(* IEC 61131-3 sources: plc-st-coding-agent/progress/evidence/f14_v10_full_20261113/jobs/codex_minimax-m27, 188 files *)

(* ---- self-hard-03.candidate_01.st ---- *)
(* ENGINEERING_CONTRACT
| Output/State    | Activation        | Retention         | Explicit Reset | Scan Priority | Units/Boundaries |
|-----------------|-------------------|-------------------|----------------|---------------|------------------|
| count           | Computed each scan| Maintained        | None           | After ops     | 0..8 integer     |
| full            | count=8           | Held until count<8| None           | With count    | BOOL             |
| empty           | count=0           | Held until count>0| None           | With count    | BOOL             |
| head            | fifo[1] or 0      | Held on empty     | None           | After ops     | INT              |
| fifo[1..count]  | Compacted each scan| Retained         | None           | After ops     | ARRAY[1..8] INT  |

PUB001: pushEn (rising edge trigger)
PUB002: pushItem (INT payload)
PUB003: popEn (rising edge trigger)
PUB004: fifo INOUT ARRAY[1..8] INT, caller-bound, read-write during scan
PUB005: count = length 0..8
PUB006: full <-> count=8
PUB007: empty <-> count=0
PUB008: head = fifo[1] when !empty else 0
PUB009: pop on rising(popEn) executes first if count>0
PUB010: push on rising(pushEn) executes second if count<8
PUB011: same-scan full+pop+push: pop frees slot then push appends
PUB012: same-scan empty+pop+push: only push adds item
PUB013: fifo[1..count] compact, fifo[1]=head when !empty
PUB014: undefined fifo[count+1..8]
PUB015: initial count=0, empty=TRUE, fifo[1..8] undefined
PUB016: rising edge = prev=FALSE AND cur=TRUE
PUB017: sustained press does not repeat (edge-only)
PUB018: R_TRIG used for edge memory
PUB019: scan-order: detect edges, execute pop, execute push, compute outputs
PUB020: CONTRACT_RULES []

Function Block FB
VAR_INPUT
    pushEn : BOOL;
    pushItem : INT;
    popEn : BOOL;
END_VAR
VAR_IN_OUT
    fifo : ARRAY[1..8] OF INT;
END_VAR
VAR_OUTPUT
    count : INT := 0;
    full : BOOL := FALSE;
    empty : BOOL := TRUE;
    head : INT := 0;
END_VAR
VAR
    pushTrig : R_TRIG;
    popTrig : R_TRIG;
END_VAR

pushTrig(CLK := pushEn);
popTrig(CLK := popEn);

IF popTrig.Q AND count > 0 THEN
    FOR i := 1 TO count - 1 DO
        fifo[i] := fifo[i + 1];
    END_FOR;
    count := count - 1;
END_IF;

IF pushTrig.Q AND count < 8 THEN
    count := count + 1;
    fifo[count] := pushItem;
END_IF;

full := (count = 8);
empty := (count = 0);
head := 0;
IF NOT empty THEN
    head := fifo[1];
END_IF;

END_FUNCTION_BLOCK

(* ---- self-hard-03.raw_candidate_01.st ---- *)
(* ENGINEERING_CONTRACT
| Output/State    | Activation        | Retention         | Explicit Reset | Scan Priority | Units/Boundaries |
|-----------------|-------------------|-------------------|----------------|---------------|------------------|
| count           | Computed each scan| Maintained        | None           | After ops     | 0..8 integer     |
| full            | count=8           | Held until count<8| None           | With count    | BOOL             |
| empty           | count=0           | Held until count>0| None           | With count    | BOOL             |
| head            | fifo[1] or 0      | Held on empty     | None           | After ops     | INT              |
| fifo[1..count]  | Compacted each scan| Retained         | None           | After ops     | ARRAY[1..8] INT  |

PUB001: pushEn (rising edge trigger)
PUB002: pushItem (INT payload)
PUB003: popEn (rising edge trigger)
PUB004: fifo INOUT ARRAY[1..8] INT, caller-bound, read-write during scan
PUB005: count = length 0..8
PUB006: full <-> count=8
PUB007: empty <-> count=0
PUB008: head = fifo[1] when !empty else 0
PUB009: pop on rising(popEn) executes first if count>0
PUB010: push on rising(pushEn) executes second if count<8
PUB011: same-scan full+pop+push: pop frees slot then push appends
PUB012: same-scan empty+pop+push: only push adds item
PUB013: fifo[1..count] compact, fifo[1]=head when !empty
PUB014: undefined fifo[count+1..8]
PUB015: initial count=0, empty=TRUE, fifo[1..8] undefined
PUB016: rising edge = prev=FALSE AND cur=TRUE
PUB017: sustained press does not repeat (edge-only)
PUB018: R_TRIG used for edge memory
PUB019: scan-order: detect edges, execute pop, execute push, compute outputs
PUB020: CONTRACT_RULES []

Function Block FB
VAR_INPUT
    pushEn : BOOL;
    pushItem : INT;
    popEn : BOOL;
END_VAR
VAR_IN_OUT
    fifo : ARRAY[1..8] OF INT;
END_VAR
VAR_OUTPUT
    count : INT := 0;
    full : BOOL := FALSE;
    empty : BOOL := TRUE;
    head : INT := 0;
END_VAR
VAR
    pushTrig : R_TRIG;
    popTrig : R_TRIG;
END_VAR

pushTrig(CLK := pushEn);
popTrig(CLK := popEn);

IF popTrig.Q AND count > 0 THEN
    FOR i := 1 TO count - 1 DO
        fifo[i] := fifo[i + 1];
    END_FOR;
    count := count - 1;
END_IF;

IF pushTrig.Q AND count < 8 THEN
    count := count + 1;
    fifo[count] := pushItem;
END_IF;

full := (count = 8);
empty := (count = 0);
head := 0;
IF NOT empty THEN
    head := fifo[1];
END_IF;

END_FUNCTION_BLOCK

(* ---- public-easy-01.candidate_01.st ---- *)
(* ENGINEERING_CONTRACT *)
(*
State  | Activation                    | Retention               | Reset/Deactivation              | Same-scan Priority | Units/Boundaries
-------|-------------------------------|-------------------------|----------------------------------|--------------------|------------------
IDLE   | bottleSensor = TRUE           | All outputs = FALSE     | None (waiting for bottle)        | -                  | edge-triggered on bottle arrival
CLEAN  | State=IDLE & bottleSensor     | Pump_Motor = TRUE       | cleaningConfirmButton = TRUE    | same-scan          | pump latches until confirmed
FILL   | cleaningConfirmButton=TRUE    | Filling_Valve = TRUE    | fillingConfirmButton = TRUE     | same-scan          | valve latches until confirmed
CAP    | fillingConfirmButton=TRUE     | Capping_Machine = TRUE  | cappingConfirmButton = TRUE     | same-scan          | machine latches until confirmed
PACK   | cappingConfirmButton=TRUE     | Packing_Machine = TRUE  | packingConfirmButton = TRUE     | same-scan          | machine latches until confirmed
DONE   | packingConfirmButton=TRUE     | Completion_Light=TRUE   | finishedButton = TRUE           | same-scan          | light stays on until reset
*)

(* CONTRACT_RULES [] *)

FUNCTION_BLOCK FillingLineControl
VAR
    State : UINT := 0; // 0=IDLE, 1=CLEAN, 2=FILL, 3=CAP, 4=PACK, 5=DONE
END_VAR

// State machine logic
CASE State OF
    0: // IDLE - Waiting for bottle
        Pump_Motor := FALSE;
        Filling_Valve := FALSE;
        Capping_Machine := FALSE;
        Packing_Machine := FALSE;
        Completion_Light := FALSE;

        IF bottleSensor THEN
            State := 1;
        END_IF;

    1: // CLEAN - Cleaning pump running
        Pump_Motor := TRUE;
        Filling_Valve := FALSE;
        Capping_Machine := FALSE;
        Packing_Machine := FALSE;
        Completion_Light := FALSE;

        IF cleaningConfirmButton THEN
            State := 2;
        END_IF;

    2: // FILL - Filling valve open
        Pump_Motor := FALSE;
        Filling_Valve := TRUE;
        Capping_Machine := FALSE;
        Packing_Machine := FALSE;
        Completion_Light := FALSE;

        IF fillingConfirmButton THEN
            State := 3;
        END_IF;

    3: // CAP - Capping machine running
        Pump_Motor := FALSE;
        Filling_Valve := FALSE;
        Capping_Machine := TRUE;
        Packing_Machine := FALSE;
        Completion_Light := FALSE;

        IF cappingConfirmButton THEN
            State := 4;
        END_IF;

    4: // PACK - Packing machine running
        Pump_Motor := FALSE;
        Filling_Valve := FALSE;
        Capping_Machine := FALSE;
        Packing_Machine := TRUE;
        Completion_Light := FALSE;

        IF packingConfirmButton THEN
            State := 5;
        END_IF;

    5: // DONE - Packaging complete, waiting for pickup
        Pump_Motor := FALSE;
        Filling_Valve := FALSE;
        Capping_Machine := FALSE;
        Packing_Machine := FALSE;
        Completion_Light := TRUE;

        IF finishedButton THEN
            State := 0;
        END_IF;

END_CASE;

END_FUNCTION_BLOCK

(* ---- public-easy-01.candidate_02.st ---- *)
(* ENGINEERING_CONTRACT *)
(*
State  | Activation                    | Retention               | Reset/Deactivation              | Same-scan Priority | Units/Boundaries
-------|-------------------------------|-------------------------|----------------------------------|--------------------|------------------
IDLE   | bottleSensor = TRUE           | All outputs = FALSE     | None (waiting for bottle)        | -                  | edge-triggered on bottle arrival
CLEAN  | State=IDLE & bottleSensor     | Pump_Motor = TRUE       | cleaningConfirmButton = TRUE    | same-scan          | pump latches until confirmed
FILL   | cleaningConfirmButton=TRUE    | Filling_Valve = TRUE    | fillingConfirmButton = TRUE     | same-scan          | valve latches until confirmed
CAP    | fillingConfirmButton=TRUE     | Capping_Machine = TRUE  | cappingConfirmButton = TRUE     | same-scan          | machine latches until confirmed
PACK   | cappingConfirmButton=TRUE     | Packing_Machine = TRUE  | packingConfirmButton = TRUE     | same-scan          | machine latches until confirmed
DONE   | packingConfirmButton=TRUE     | Completion_Light=TRUE   | finishedButton = TRUE           | same-scan          | light stays on until reset
*)

(* CONTRACT_RULES [] *)

FUNCTION_BLOCK FillingLineControl
VAR_INPUT
    bottleSensor : BOOL;
    cleaningConfirmButton : BOOL;
    fillingConfirmButton : BOOL;
    cappingConfirmButton : BOOL;
    packingConfirmButton : BOOL;
    finishedButton : BOOL;
END_VAR

VAR_OUTPUT
    Pump_Motor : BOOL;
    Filling_Valve : BOOL;
    Capping_Machine : BOOL;
    Packing_Machine : BOOL;
    Completion_Light : BOOL;
END_VAR

VAR
    State : UINT := 0;
END_VAR

CASE State OF
    0:
        Pump_Motor := FALSE;
        Filling_Valve := FALSE;
        Capping_Machine := FALSE;
        Packing_Machine := FALSE;
        Completion_Light := FALSE;

        IF bottleSensor THEN
            State := 1;
        END_IF;

    1:
        Pump_Motor := TRUE;
        Filling_Valve := FALSE;
        Capping_Machine := FALSE;
        Packing_Machine := FALSE;
        Completion_Light := FALSE;

        IF cleaningConfirmButton THEN
            State := 2;
        END_IF;

    2:
        Pump_Motor := FALSE;
        Filling_Valve := TRUE;
        Capping_Machine := FALSE;
        Packing_Machine := FALSE;
        Completion_Light := FALSE;

        IF fillingConfirmButton THEN
            State := 3;
        END_IF;

    3:
        Pump_Motor := FALSE;
        Filling_Valve := FALSE;
        Capping_Machine := TRUE;
        Packing_Machine := FALSE;
        Completion_Light := FALSE;

        IF cappingConfirmButton THEN
            State := 4;
        END_IF;

    4:
        Pump_Motor := FALSE;
        Filling_Valve := FALSE;
        Capping_Machine := FALSE;
        Packing_Machine := TRUE;
        Completion_Light := FALSE;

        IF packingConfirmButton THEN
            State := 5;
        END_IF;

    5:
        Pump_Motor := FALSE;
        Filling_Valve := FALSE;
        Capping_Machine := FALSE;
        Packing_Machine := FALSE;
        Completion_Light := TRUE;

        IF finishedButton THEN
            State := 0;
        END_IF;

END_CASE;

END_FUNCTION_BLOCK

(* ---- public-easy-01.candidate_03.st ---- *)
Looking at the test failures, I can see the issue: in the original code, when a state transition occurs (e.g., from state 0 to 1 when bottleSensor is true), the CASE statement continues executing remaining assignments in that branch based on the **new** state value, causing outputs to reflect the next state rather than the triggering state.

For example, when bottleSensor=TRUE in state 0, State becomes 1, but then assignments for state 1 execute in the same branch, setting Pump_Motor=TRUE. But for tc-02 (single scan, bottleSensor=TRUE), the expected output should be Pump_Motor=TRUE... wait, the checkpoint shows Pump_Motor=FALSE.

Let me trace more carefully. The issue is that outputs are computed **during** the transition case branch, reading the **updated** State value. The fix is to separate transition computation from output computation.

(* ENGINEERING_CONTRACT *)
(*
State  | Activation                    | Retention               | Reset/Deactivation              | Same-scan Priority | Units/Boundaries
-------|-------------------------------|-------------------------|----------------------------------|--------------------|------------------
IDLE   | bottleSensor = TRUE           | All outputs = FALSE     | None (waiting for bottle)        | -                  | edge-triggered on bottle arrival
CLEAN  | State=IDLE & bottleSensor     | Pump_Motor = TRUE       | cleaningConfirmButton = TRUE    | same-scan          | pump latches until confirmed
FILL   | cleaningConfirmButton=TRUE    | Filling_Valve = TRUE    | fillingConfirmButton = TRUE     | same-scan          | valve latches until confirmed
CAP    | fillingConfirmButton=TRUE     | Capping_Machine = TRUE  | cappingConfirmButton = TRUE     | same-scan          | machine latches until confirmed
PACK   | cappingConfirmButton=TRUE     | Packing_Machine = TRUE  | packingConfirmButton = TRUE     | same-scan          | machine latches until confirmed
DONE   | packingConfirmButton=TRUE     | Completion_Light=TRUE   | finishedButton = TRUE           | same-scan          | light stays on until reset
*)

(* CONTRACT_RULES [] *)

FUNCTION_BLOCK FillingLineControl
VAR_INPUT
    bottleSensor : BOOL;
    cleaningConfirmButton : BOOL;
    fillingConfirmButton : BOOL;
    cappingConfirmButton : BOOL;
    packingConfirmButton : BOOL;
    finishedButton : BOOL;
END_VAR

VAR_OUTPUT
    Pump_Motor : BOOL;
    Filling_Valve : BOOL;
    Capping_Machine : BOOL;
    Packing_Machine : BOOL;
    Completion_Light : BOOL;
END_VAR

VAR
    State : UINT := 0;
    tmp_nextState : UINT := 0;
END_VAR

CASE State OF
    0:
        tmp_nextState := 0;
        IF bottleSensor THEN
            tmp_nextState := 1;
        END_IF;

    1:
        tmp_nextState := 1;
        IF cleaningConfirmButton THEN
            tmp_nextState := 2;
        END_IF;

    2:
        tmp_nextState := 2;
        IF fillingConfirmButton THEN
            tmp_nextState := 3;
        END_IF;

    3:
        tmp_nextState := 3;
        IF cappingConfirmButton THEN
            tmp_nextState := 4;
        END_IF;

    4:
        tmp_nextState := 4;
        IF packingConfirmButton THEN
            tmp_nextState := 5;
        END_IF;

    5:
        tmp_nextState := 5;
        IF finishedButton THEN
            tmp_nextState := 0;
        END_IF;
END_CASE;

State := tmp_nextState;

CASE State OF
    0:
        Pump_Motor := FALSE;
        Filling_Valve := FALSE;
        Capping_Machine := FALSE;
        Packing_Machine := FALSE;
        Completion_Light := FALSE;

    1:
        Pump_Motor := TRUE;
        Filling_Valve := FALSE;
        Capping_Machine := FALSE;
        Packing_Machine := FALSE;
        Completion_Light := FALSE;

    2:
        Pump_Motor := FALSE;
        Filling_Valve := TRUE;
        Capping_Machine := FALSE;
        Packing_Machine := FALSE;
        Completion_Light := FALSE;

    3:
        Pump_Motor := FALSE;
        Filling_Valve := FALSE;
        Capping_Machine := TRUE;
        Packing_Machine := FALSE;
        Completion_Light := FALSE;

    4:
        Pump_Motor := FALSE;
        Filling_Valve := FALSE;
        Capping_Machine := FALSE;
        Packing_Machine := TRUE;
        Completion_Light := FALSE;

    5:
        Pump_Motor := FALSE;
        Filling_Valve := FALSE;
        Capping_Machine := FALSE;
        Packing_Machine := FALSE;
        Completion_Light := TRUE;

END_CASE;

END_FUNCTION_BLOCK

(* ---- public-easy-01.raw_candidate_01.st ---- *)
(* ENGINEERING_CONTRACT *)
(*
State  | Activation                    | Retention               | Reset/Deactivation              | Same-scan Priority | Units/Boundaries
-------|-------------------------------|-------------------------|----------------------------------|--------------------|------------------
IDLE   | bottleSensor = TRUE           | All outputs = FALSE     | None (waiting for bottle)        | -                  | edge-triggered on bottle arrival
CLEAN  | State=IDLE & bottleSensor     | Pump_Motor = TRUE       | cleaningConfirmButton = TRUE    | same-scan          | pump latches until confirmed
FILL   | cleaningConfirmButton=TRUE    | Filling_Valve = TRUE    | fillingConfirmButton = TRUE     | same-scan          | valve latches until confirmed
CAP    | fillingConfirmButton=TRUE     | Capping_Machine = TRUE  | cappingConfirmButton = TRUE     | same-scan          | machine latches until confirmed
PACK   | cappingConfirmButton=TRUE     | Packing_Machine = TRUE  | packingConfirmButton = TRUE     | same-scan          | machine latches until confirmed
DONE   | packingConfirmButton=TRUE     | Completion_Light=TRUE   | finishedButton = TRUE           | same-scan          | light stays on until reset
*)

(* CONTRACT_RULES [] *)

FUNCTION_BLOCK FillingLineControl
VAR
    State : UINT := 0; // 0=IDLE, 1=CLEAN, 2=FILL, 3=CAP, 4=PACK, 5=DONE
END_VAR

// State machine logic
CASE State OF
    0: // IDLE - Waiting for bottle
        Pump_Motor := FALSE;
        Filling_Valve := FALSE;
        Capping_Machine := FALSE;
        Packing_Machine := FALSE;
        Completion_Light := FALSE;

        IF bottleSensor THEN
            State := 1;
        END_IF

    1: // CLEAN - Cleaning pump running
        Pump_Motor := TRUE;
        Filling_Valve := FALSE;
        Capping_Machine := FALSE;
        Packing_Machine := FALSE;
        Completion_Light := FALSE;

        IF cleaningConfirmButton THEN
            State := 2;
        END_IF

    2: // FILL - Filling valve open
        Pump_Motor := FALSE;
        Filling_Valve := TRUE;
        Capping_Machine := FALSE;
        Packing_Machine := FALSE;
        Completion_Light := FALSE;

        IF fillingConfirmButton THEN
            State := 3;
        END_IF

    3: // CAP - Capping machine running
        Pump_Motor := FALSE;
        Filling_Valve := FALSE;
        Capping_Machine := TRUE;
        Packing_Machine := FALSE;
        Completion_Light := FALSE;

        IF cappingConfirmButton THEN
            State := 4;
        END_IF

    4: // PACK - Packing machine running
        Pump_Motor := FALSE;
        Filling_Valve := FALSE;
        Capping_Machine := FALSE;
        Packing_Machine := TRUE;
        Completion_Light := FALSE;

        IF packingConfirmButton THEN
            State := 5;
        END_IF

    5: // DONE - Packaging complete, waiting for pickup
        Pump_Motor := FALSE;
        Filling_Valve := FALSE;
        Capping_Machine := FALSE;
        Packing_Machine := FALSE;
        Completion_Light := TRUE;

        IF finishedButton THEN
            State := 0;
        END_IF

END_CASE;

END_FUNCTION_BLOCK

(* ---- public-easy-01.raw_candidate_02.st ---- *)
(* ENGINEERING_CONTRACT *)
(*
State  | Activation                    | Retention               | Reset/Deactivation              | Same-scan Priority | Units/Boundaries
-------|-------------------------------|-------------------------|----------------------------------|--------------------|------------------
IDLE   | bottleSensor = TRUE           | All outputs = FALSE     | None (waiting for bottle)        | -                  | edge-triggered on bottle arrival
CLEAN  | State=IDLE & bottleSensor     | Pump_Motor = TRUE       | cleaningConfirmButton = TRUE    | same-scan          | pump latches until confirmed
FILL   | cleaningConfirmButton=TRUE    | Filling_Valve = TRUE    | fillingConfirmButton = TRUE     | same-scan          | valve latches until confirmed
CAP    | fillingConfirmButton=TRUE     | Capping_Machine = TRUE  | cappingConfirmButton = TRUE     | same-scan          | machine latches until confirmed
PACK   | cappingConfirmButton=TRUE     | Packing_Machine = TRUE  | packingConfirmButton = TRUE     | same-scan          | machine latches until confirmed
DONE   | packingConfirmButton=TRUE     | Completion_Light=TRUE   | finishedButton = TRUE           | same-scan          | light stays on until reset
*)

(* CONTRACT_RULES [] *)

FUNCTION_BLOCK FillingLineControl
VAR_INPUT
    bottleSensor : BOOL;
    cleaningConfirmButton : BOOL;
    fillingConfirmButton : BOOL;
    cappingConfirmButton : BOOL;
    packingConfirmButton : BOOL;
    finishedButton : BOOL;
END_VAR

VAR_OUTPUT
    Pump_Motor : BOOL;
    Filling_Valve : BOOL;
    Capping_Machine : BOOL;
    Packing_Machine : BOOL;
    Completion_Light : BOOL;
END_VAR

VAR
    State : UINT := 0;
END_VAR

CASE State OF
    0:
        Pump_Motor := FALSE;
        Filling_Valve := FALSE;
        Capping_Machine := FALSE;
        Packing_Machine := FALSE;
        Completion_Light := FALSE;

        IF bottleSensor THEN
            State := 1;
        END_IF;

    1:
        Pump_Motor := TRUE;
        Filling_Valve := FALSE;
        Capping_Machine := FALSE;
        Packing_Machine := FALSE;
        Completion_Light := FALSE;

        IF cleaningConfirmButton THEN
            State := 2;
        END_IF;

    2:
        Pump_Motor := FALSE;
        Filling_Valve := TRUE;
        Capping_Machine := FALSE;
        Packing_Machine := FALSE;
        Completion_Light := FALSE;

        IF fillingConfirmButton THEN
            State := 3;
        END_IF;

    3:
        Pump_Motor := FALSE;
        Filling_Valve := FALSE;
        Capping_Machine := TRUE;
        Packing_Machine := FALSE;
        Completion_Light := FALSE;

        IF cappingConfirmButton THEN
            State := 4;
        END_IF;

    4:
        Pump_Motor := FALSE;
        Filling_Valve := FALSE;
        Capping_Machine := FALSE;
        Packing_Machine := TRUE;
        Completion_Light := FALSE;

        IF packingConfirmButton THEN
            State := 5;
        END_IF;

    5:
        Pump_Motor := FALSE;
        Filling_Valve := FALSE;
        Capping_Machine := FALSE;
        Packing_Machine := FALSE;
        Completion_Light := TRUE;

        IF finishedButton THEN
            State := 0;
        END_IF;

END_CASE;

END_FUNCTION_BLOCK

(* ---- public-easy-01.raw_candidate_03.st ---- *)
Looking at the test failures, I can see the issue: in the original code, when a state transition occurs (e.g., from state 0 to 1 when bottleSensor is true), the CASE statement continues executing remaining assignments in that branch based on the **new** state value, causing outputs to reflect the next state rather than the triggering state.

For example, when bottleSensor=TRUE in state 0, State becomes 1, but then assignments for state 1 execute in the same branch, setting Pump_Motor=TRUE. But for tc-02 (single scan, bottleSensor=TRUE), the expected output should be Pump_Motor=TRUE... wait, the checkpoint shows Pump_Motor=FALSE.

Let me trace more carefully. The issue is that outputs are computed **during** the transition case branch, reading the **updated** State value. The fix is to separate transition computation from output computation.

(* ENGINEERING_CONTRACT *)
(*
State  | Activation                    | Retention               | Reset/Deactivation              | Same-scan Priority | Units/Boundaries
-------|-------------------------------|-------------------------|----------------------------------|--------------------|------------------
IDLE   | bottleSensor = TRUE           | All outputs = FALSE     | None (waiting for bottle)        | -                  | edge-triggered on bottle arrival
CLEAN  | State=IDLE & bottleSensor     | Pump_Motor = TRUE       | cleaningConfirmButton = TRUE    | same-scan          | pump latches until confirmed
FILL   | cleaningConfirmButton=TRUE    | Filling_Valve = TRUE    | fillingConfirmButton = TRUE     | same-scan          | valve latches until confirmed
CAP    | fillingConfirmButton=TRUE     | Capping_Machine = TRUE  | cappingConfirmButton = TRUE     | same-scan          | machine latches until confirmed
PACK   | cappingConfirmButton=TRUE     | Packing_Machine = TRUE  | packingConfirmButton = TRUE     | same-scan          | machine latches until confirmed
DONE   | packingConfirmButton=TRUE     | Completion_Light=TRUE   | finishedButton = TRUE           | same-scan          | light stays on until reset
*)

(* CONTRACT_RULES [] *)

FUNCTION_BLOCK FillingLineControl
VAR_INPUT
    bottleSensor : BOOL;
    cleaningConfirmButton : BOOL;
    fillingConfirmButton : BOOL;
    cappingConfirmButton : BOOL;
    packingConfirmButton : BOOL;
    finishedButton : BOOL;
END_VAR

VAR_OUTPUT
    Pump_Motor : BOOL;
    Filling_Valve : BOOL;
    Capping_Machine : BOOL;
    Packing_Machine : BOOL;
    Completion_Light : BOOL;
END_VAR

VAR
    State : UINT := 0;
    tmp_nextState : UINT := 0;
END_VAR

CASE State OF
    0:
        tmp_nextState := 0;
        IF bottleSensor THEN
            tmp_nextState := 1;
        END_IF;

    1:
        tmp_nextState := 1;
        IF cleaningConfirmButton THEN
            tmp_nextState := 2;
        END_IF;

    2:
        tmp_nextState := 2;
        IF fillingConfirmButton THEN
            tmp_nextState := 3;
        END_IF;

    3:
        tmp_nextState := 3;
        IF cappingConfirmButton THEN
            tmp_nextState := 4;
        END_IF;

    4:
        tmp_nextState := 4;
        IF packingConfirmButton THEN
            tmp_nextState := 5;
        END_IF;

    5:
        tmp_nextState := 5;
        IF finishedButton THEN
            tmp_nextState := 0;
        END_IF;
END_CASE;

State := tmp_nextState;

CASE State OF
    0:
        Pump_Motor := FALSE;
        Filling_Valve := FALSE;
        Capping_Machine := FALSE;
        Packing_Machine := FALSE;
        Completion_Light := FALSE;

    1:
        Pump_Motor := TRUE;
        Filling_Valve := FALSE;
        Capping_Machine := FALSE;
        Packing_Machine := FALSE;
        Completion_Light := FALSE;

    2:
        Pump_Motor := FALSE;
        Filling_Valve := TRUE;
        Capping_Machine := FALSE;
        Packing_Machine := FALSE;
        Completion_Light := FALSE;

    3:
        Pump_Motor := FALSE;
        Filling_Valve := FALSE;
        Capping_Machine := TRUE;
        Packing_Machine := FALSE;
        Completion_Light := FALSE;

    4:
        Pump_Motor := FALSE;
        Filling_Valve := FALSE;
        Capping_Machine := FALSE;
        Packing_Machine := TRUE;
        Completion_Light := FALSE;

    5:
        Pump_Motor := FALSE;
        Filling_Valve := FALSE;
        Capping_Machine := FALSE;
        Packing_Machine := FALSE;
        Completion_Light := TRUE;

END_CASE;

END_FUNCTION_BLOCK

(* ---- public-easy-02.candidate_01.st ---- *)
FUNCTION_BLOCK FB_DualWordEdgeDetector
VAR_INPUT
END_VAR
VAR_OUTPUT
    hasChanged     : BOOL  := FALSE;
    hasRisingEdges : BOOL  := FALSE;
    risingBits     : DWORD := 0;
    noOfRisingBits : USINT := 0;
    hasFallingEdges: BOOL  := FALSE;
    fallingBits    : DWORD := 0;
    noOfFallingBits: USINT := 0;
END_VAR
VAR
    previousValue : DWORD := 0;
    tmpXorMask    : DWORD;
    tmpRising     : DWORD;
    tmpFalling    : DWORD;
    tmpIdx        : USINT;
END_VAR
VAR_TEMP
END_VAR
(*
ENGINEERING_CONTRACT
===================
PUB001: Dual-word edge detection every scan cycle
-----------------------------------------------
Output/State    | Activation           | Retention    | Reset        | Priority     | Units/Boundary
----------------|----------------------|--------------|--------------|--------------|-----------------
hasChanged      | value <> prev        | per scan     | auto-clear   | same-scan    | BOOL
risingBits      | cur=1 AND prev=0     | per scan     | auto-clear   | same-scan    | DWORD mask
noOfRisingBits  | count(risingBits)    | per scan     | auto-clear   | same-scan    | 0..32
hasFallingEdges | fallingBits <> 0     | per scan     | auto-clear   | same-scan    | BOOL
fallingBits     | cur=0 AND prev=1     | per scan     | auto-clear   | same-scan    | DWORD mask
noOfFallingBits | count(fallingBits)   | per scan     | auto-clear   | same-scan    | 0..32
previousValue   | hold across scans    | retained     | no reset     | same-scan    | DWORD

Same-scan behavior: All outputs derived from (value, previousValue) on each invocation.
No edge-only triggers or external resets are specified.
*)
tmpXorMask := value XOR previousValue;
tmpRising  := tmpXorMask AND value;
tmpFalling := tmpXorMask AND previousValue;

hasChanged      := (value <> previousValue);
hasRisingEdges  := (tmpRising <> 0);
hasFallingEdges := (tmpFalling <> 0);
risingBits      := tmpRising;
fallingBits     := tmpFalling;

noOfRisingBits  := 0;
noOfFallingBits := 0;
FOR tmpIdx := 0 TO 31 DO
    IF (SHR(risingBits, TO_UINT(tmpIdx)) AND 1) = 1 THEN
        noOfRisingBits := noOfRisingBits + 1;
    END_IF;
    IF (SHR(fallingBits, TO_UINT(tmpIdx)) AND 1) = 1 THEN
        noOfFallingBits := noOfFallingBits + 1;
    END_IF;
END_FOR;

previousValue := value;
END_FUNCTION_BLOCK
(* CONTRACT_RULES [] *)

(* ---- public-easy-02.raw_candidate_01.st ---- *)
FUNCTION_BLOCK FB_DualWordEdgeDetector
VAR_INPUT
END_VAR
VAR_OUTPUT
    hasChanged     : BOOL  := FALSE;
    hasRisingEdges : BOOL  := FALSE;
    risingBits     : DWORD := 0;
    noOfRisingBits : USINT := 0;
    hasFallingEdges: BOOL  := FALSE;
    fallingBits    : DWORD := 0;
    noOfFallingBits: USINT := 0;
END_VAR
VAR
    previousValue : DWORD := 0;
    tmpXorMask    : DWORD;
    tmpRising     : DWORD;
    tmpFalling    : DWORD;
    tmpIdx        : USINT;
END_VAR
VAR_TEMP
END_VAR
(*
ENGINEERING_CONTRACT
===================
PUB001: Dual-word edge detection every scan cycle
-----------------------------------------------
Output/State    | Activation           | Retention    | Reset        | Priority     | Units/Boundary
----------------|----------------------|--------------|--------------|--------------|-----------------
hasChanged      | value <> prev        | per scan     | auto-clear   | same-scan    | BOOL
risingBits      | cur=1 AND prev=0     | per scan     | auto-clear   | same-scan    | DWORD mask
noOfRisingBits  | count(risingBits)    | per scan     | auto-clear   | same-scan    | 0..32
hasFallingEdges | fallingBits <> 0     | per scan     | auto-clear   | same-scan    | BOOL
fallingBits     | cur=0 AND prev=1     | per scan     | auto-clear   | same-scan    | DWORD mask
noOfFallingBits | count(fallingBits)   | per scan     | auto-clear   | same-scan    | 0..32
previousValue   | hold across scans    | retained     | no reset     | same-scan    | DWORD

Same-scan behavior: All outputs derived from (value, previousValue) on each invocation.
No edge-only triggers or external resets are specified.
*)
tmpXorMask := value XOR previousValue;
tmpRising  := tmpXorMask AND value;
tmpFalling := tmpXorMask AND previousValue;

hasChanged      := (value <> previousValue);
hasRisingEdges  := (tmpRising <> 0);
hasFallingEdges := (tmpFalling <> 0);
risingBits      := tmpRising;
fallingBits     := tmpFalling;

noOfRisingBits  := 0;
noOfFallingBits := 0;
FOR tmpIdx := 0 TO 31 DO
    IF (SHR(risingBits, TO_UINT(tmpIdx)) AND 1) = 1 THEN
        noOfRisingBits := noOfRisingBits + 1;
    END_IF
    IF (SHR(fallingBits, TO_UINT(tmpIdx)) AND 1) = 1 THEN
        noOfFallingBits := noOfFallingBits + 1;
    END_IF
END_FOR

previousValue := value;
END_FUNCTION_BLOCK
(* CONTRACT_RULES [] *)

(* ---- public-easy-03.candidate_01.st ---- *)
FUNCTION_BLOCK AlarmWithHysteresis
VAR_OUTPUT
    hiAlarm : BOOL := FALSE;
    loAlarm : BOOL := FALSE;
    error   : BOOL := FALSE;
    status  : WORD := 16#0000;
END_VAR
VAR_INPUT
    Value      : REAL;
    hiLevel    : REAL;
    loLevel    : REAL;
    hystWindow : REAL;
END_VAR

// ENGINEERING_CONTRACT
// State retention: hiAlarm and loAlarm hold state across scans (level-triggered behavior)
// PUB001: hiAlarm activates at Value > hiLevel, deactivates at Value < hiLevel - hystWindow
// PUB002: loAlarm activates at Value < loLevel, deactivates at Value > loLevel + hystWindow
// PUB003: error=TRUE and status=16#8001 if loLevel >= hiLevel (checked first)
// PUB004: error=TRUE and status=16#8002 if hystWindow >= (hiLevel - loLevel)
// PUB005-PUB007: On error, set error=TRUE with status, exit without changing alarm outputs
// Same-scan priority: Error checks first, then hiAlarm, then loAlarm evaluation
// Units/boundaries: REAL comparison; error codes 16#8001, 16#8002; default status=16#0000

// CONTRACT_RULES: []
// No unconditional Boolean output latches; alarms are level-triggered based on current Value

// Error checking - highest priority
IF loLevel >= hiLevel THEN
    error := TRUE;
    status := 16#8001;
    RETURN;
END_IF;

IF hystWindow >= (hiLevel - loLevel) THEN
    error := TRUE;
    status := 16#8002;
    RETURN;
END_IF;

// No error; evaluate alarms based on current Value
error := FALSE;
status := 16#0000;

IF Value > hiLevel THEN
    hiAlarm := TRUE;
ELSIF Value < (hiLevel - hystWindow) THEN
    hiAlarm := FALSE;
END_IF;

IF Value < loLevel THEN
    loAlarm := TRUE;
ELSIF Value > (loLevel + hystWindow) THEN
    loAlarm := FALSE;
END_IF;

END_FUNCTION_BLOCK

(* ---- public-easy-03.raw_candidate_01.st ---- *)
FUNCTION_BLOCK AlarmWithHysteresis
VAR_OUTPUT
    hiAlarm : BOOL := FALSE;
    loAlarm : BOOL := FALSE;
    error   : BOOL := FALSE;
    status  : WORD := 16#0000;
END_VAR
VAR_INPUT
    Value      : REAL;
    hiLevel    : REAL;
    loLevel    : REAL;
    hystWindow : REAL;
END_VAR

// ENGINEERING_CONTRACT
// State retention: hiAlarm and loAlarm hold state across scans (level-triggered behavior)
// PUB001: hiAlarm activates at Value > hiLevel, deactivates at Value < hiLevel - hystWindow
// PUB002: loAlarm activates at Value < loLevel, deactivates at Value > loLevel + hystWindow
// PUB003: error=TRUE and status=16#8001 if loLevel >= hiLevel (checked first)
// PUB004: error=TRUE and status=16#8002 if hystWindow >= (hiLevel - loLevel)
// PUB005-PUB007: On error, set error=TRUE with status, exit without changing alarm outputs
// Same-scan priority: Error checks first, then hiAlarm, then loAlarm evaluation
// Units/boundaries: REAL comparison; error codes 16#8001, 16#8002; default status=16#0000

// CONTRACT_RULES: []
// No unconditional Boolean output latches; alarms are level-triggered based on current Value

// Error checking - highest priority
IF loLevel >= hiLevel THEN
    error := TRUE;
    status := 16#8001;
    RETURN;
END_IF

IF hystWindow >= (hiLevel - loLevel) THEN
    error := TRUE;
    status := 16#8002;
    RETURN;
END_IF

// No error; evaluate alarms based on current Value
error := FALSE;
status := 16#0000;

IF Value > hiLevel THEN
    hiAlarm := TRUE;
ELSIF Value < (hiLevel - hystWindow) THEN
    hiAlarm := FALSE;
END_IF;

IF Value < loLevel THEN
    loAlarm := TRUE;
ELSIF Value > (loLevel + hystWindow) THEN
    loAlarm := FALSE;
END_IF;

END_FUNCTION_BLOCK

(* ---- public-easy-04.candidate_01.st ---- *)
(* ENGINEERING_CONTRACT
+------------------------------------------------------------------+
| Output/State  | Activation | Retention | Reset/Deactivation      |
+------------------------------------------------------------------+
| VFD_RUN       | TRUE when EStop=TRUE AND ViscosityValid=TRUE     |  PUB002
|               | (same-scan priority; no edge trigger)            |
+------------------------------------------------------------------+
| VFD_RUN       | Deactivates immediately when PASTE_E_STOP_NC=FALSE| PUB002
|               | or when ViscosityValid transitions to FALSE      |
+------------------------------------------------------------------+
| ViscosityValid| TRUE after VISCOSITY_OK held TRUE >= DebounceTime | PUB001
|               | Invalidated immediately when VISCOSITY_OK=FALSE  |
+------------------------------------------------------------------+
| ViscosityDebounce (TON) | Cleared on E-Stop or Viscosity=FALSE   | PUB002
+------------------------------------------------------------------+
| PUMP_RUNTIME_ACC | Accumulates LTIME += CycleTime while VFD_RUN   | PUB003
|                  | Retained when VFD_RUN=FALSE                   |
+------------------------------------------------------------------+
| PUMP_MAINT_DUE   | Set when PUMP_RUNTIME_ACC >= 500 hours         | PUB004
|                  | Informational only; no effect on VFD_RUN      |
+------------------------------------------------------------------+
| All outputs     | Initialize to FALSE/zero at power-up          | PUB005
+------------------------------------------------------------------+
Time boundary: 500 hours = 1,800,000,000 ms = 1,800,000,000,000 ns  PUB004
TON.Q: elapsed >= PT; first satisfying tick at ceil(DebounceTime/1ms) PUB001
CycleTime quantum: 1 ms; accumulated via LTIME nanoseconds           PUB003
+------------------------------------------------------------------+
*)
(* CONTRACT_RULES [] *)

FUNCTION_BLOCK JamPumpControl
VAR_INPUT
    VISCOSITY_OK    : BOOL;
    PASTE_E_STOP_NC : BOOL;
    DebounceTime    : TIME;
    CycleTime       : TIME;
END_VAR
VAR_OUTPUT
    VFD_RUN         : BOOL;
    PUMP_MAINT_DUE  : BOOL;
    PUMP_RUNTIME_ACC: LTIME;
END_VAR
VAR
    ViscosityValid  : BOOL := FALSE;
    ViscosityDebounce : TON;
    FirstScan       : BOOL := TRUE;
    tmpCycleNs      : LINT;
END_VAR

// Power-up initialization
IF FirstScan THEN
    VFD_RUN          := FALSE;
    PUMP_MAINT_DUE   := FALSE;
    PUMP_RUNTIME_ACC := LTIME#0s;
    FirstScan        := FALSE;
END_IF;

// Debounce state machine
ViscosityDebounce(IN  := VISCOSITY_OK AND PASTE_E_STOP_NC,
                  PT  := DebounceTime);

IF NOT VISCOSITY_OK THEN
    ViscosityValid := FALSE;
ELSIF ViscosityDebounce.Q THEN
    ViscosityValid := TRUE;
END_IF;

// VFD_RUN permissive: E-Stop OK AND viscosity condition valid
VFD_RUN := PASTE_E_STOP_NC AND ViscosityValid;

// Runtime accumulation while pump is running
IF VFD_RUN THEN
    tmpCycleNs := TO_LINT(CycleTime) * 1000000;
    PUMP_RUNTIME_ACC := PUMP_RUNTIME_ACC + TO_LTIME(tmpCycleNs);
END_IF;

// Maintenance due at 500 hours
PUMP_MAINT_DUE := PUMP_RUNTIME_ACC >= LTIME#500h;

END_FUNCTION_BLOCK

(* ---- public-easy-04.raw_candidate_01.st ---- *)
(* ENGINEERING_CONTRACT
+------------------------------------------------------------------+
| Output/State  | Activation | Retention | Reset/Deactivation      |
+------------------------------------------------------------------+
| VFD_RUN       | TRUE when EStop=TRUE AND ViscosityValid=TRUE     |  PUB002
|               | (same-scan priority; no edge trigger)            |
+------------------------------------------------------------------+
| VFD_RUN       | Deactivates immediately when PASTE_E_STOP_NC=FALSE| PUB002
|               | or when ViscosityValid transitions to FALSE      |
+------------------------------------------------------------------+
| ViscosityValid| TRUE after VISCOSITY_OK held TRUE >= DebounceTime | PUB001
|               | Invalidated immediately when VISCOSITY_OK=FALSE  |
+------------------------------------------------------------------+
| ViscosityDebounce (TON) | Cleared on E-Stop or Viscosity=FALSE   | PUB002
+------------------------------------------------------------------+
| PUMP_RUNTIME_ACC | Accumulates LTIME += CycleTime while VFD_RUN   | PUB003
|                  | Retained when VFD_RUN=FALSE                   |
+------------------------------------------------------------------+
| PUMP_MAINT_DUE   | Set when PUMP_RUNTIME_ACC >= 500 hours         | PUB004
|                  | Informational only; no effect on VFD_RUN      |
+------------------------------------------------------------------+
| All outputs     | Initialize to FALSE/zero at power-up          | PUB005
+------------------------------------------------------------------+
Time boundary: 500 hours = 1,800,000,000 ms = 1,800,000,000,000 ns  PUB004
TON.Q: elapsed >= PT; first satisfying tick at ceil(DebounceTime/1ms) PUB001
CycleTime quantum: 1 ms; accumulated via LTIME nanoseconds           PUB003
+------------------------------------------------------------------+
*)
(* CONTRACT_RULES [] *)

FUNCTION_BLOCK JamPumpControl
VAR_INPUT
    VISCOSITY_OK    : BOOL;
    PASTE_E_STOP_NC : BOOL;
    DebounceTime    : TIME;
    CycleTime       : TIME;
END_VAR
VAR_OUTPUT
    VFD_RUN         : BOOL;
    PUMP_MAINT_DUE  : BOOL;
    PUMP_RUNTIME_ACC: LTIME;
END_VAR
VAR
    ViscosityValid  : BOOL := FALSE;
    ViscosityDebounce : TON;
    FirstScan       : BOOL := TRUE;
    tmpCycleNs      : LINT;
END_VAR

// Power-up initialization
IF FirstScan THEN
    VFD_RUN          := FALSE;
    PUMP_MAINT_DUE   := FALSE;
    PUMP_RUNTIME_ACC := LTIME#0s;
    FirstScan        := FALSE;
END_IF;

// Debounce state machine
ViscosityDebounce(IN  := VISCOSITY_OK AND PASTE_E_STOP_NC,
                  PT  := DebounceTime);

IF NOT VISCOSITY_OK THEN
    ViscosityValid := FALSE;
ELSIF ViscosityDebounce.Q THEN
    ViscosityValid := TRUE;
END_IF;

// VFD_RUN permissive: E-Stop OK AND viscosity condition valid
VFD_RUN := PASTE_E_STOP_NC AND ViscosityValid;

// Runtime accumulation while pump is running
IF VFD_RUN THEN
    tmpCycleNs := TO_LINT(CycleTime) * 1000000;
    PUMP_RUNTIME_ACC := PUMP_RUNTIME_ACC + TO_LTIME(tmpCycleNs);
END_IF;

// Maintenance due at 500 hours
PUMP_MAINT_DUE := PUMP_RUNTIME_ACC >= LTIME#500h;

END_FUNCTION_BLOCK

(* ---- public-easy-05.candidate_01.st ---- *)
FUNCTION_BLOCK Weld_Gap_Alarm
(* ENGINEERING_CONTRACT
 * States: INIT(5s inhibit) | MONITOR(gap OK) | ALARM(gap debounced)
 *
 * Operator_Alert: FALSE during INIT, TRUE only when gap TRUE for >= DebounceTime
 * Weld_Soft_Start_Active: TRUE during INIT (PUB005), FALSE otherwise
 *
 * Reset/priority: E_Stop FALSE (active) >> INIT >> MONITOR/ALARM
 * - E_Stop: clears alarm, timers (PUB004)
 * - Gap FALSE: clears alarm, debounce timer (PUB003)
 * - No latching; alarm is level-driven by debounced gap
 *)
VAR_INPUT
    Gap_Exceeded   : BOOL;
    Weld_E_Stop_NC : BOOL;
    DebounceTime   : TIME;
END_VAR

VAR_OUTPUT
    Operator_Alert        : BOOL := FALSE;
    Weld_Soft_Start_Active : BOOL := TRUE;
END_VAR

VAR
    init_timer      : TON;
    debounce_timer  : TON;
    init_complete   : BOOL := FALSE;
END_VAR

    // E-Stop priority: active when Weld_E_Stop_NC = FALSE
    IF NOT Weld_E_Stop_NC THEN
        Operator_Alert         := FALSE;
        Weld_Soft_Start_Active := FALSE;
        debounce_timer(IN := FALSE);
        init_timer(IN := FALSE);
        init_complete := FALSE;
        RETURN;
    END_IF;

    // Initialization: 5-second power-up inhibition (PUB002, PUB005)
    IF NOT init_complete THEN
        init_timer(IN := TRUE, PT := T#5S);
        Weld_Soft_Start_Active := TRUE;
        Operator_Alert         := FALSE;
        debounce_timer(IN := FALSE);

        IF init_timer.Q THEN
            init_complete          := TRUE;
            Weld_Soft_Start_Active := FALSE;
            init_timer(IN := FALSE);
        END_IF;

    // Normal monitoring: debounce gap signal (PUB003)
    ELSE
        Operator_Alert := FALSE;

        IF Gap_Exceeded THEN
            debounce_timer(IN := TRUE, PT := DebounceTime);
            Operator_Alert := debounce_timer.Q;
        ELSE
            debounce_timer(IN := FALSE);
        END_IF;
    END_IF;

END_FUNCTION_BLOCK
(* CONTRACT_RULES [] *)

(* ---- public-easy-05.candidate_02.st ---- *)
FUNCTION_BLOCK Weld_Gap_Alarm
(* ENGINEERING_CONTRACT
 * States: INIT(5s inhibit) | MONITOR(gap OK) | ALARM(gap debounced)
 *
 * Operator_Alert: FALSE during INIT, TRUE only when gap TRUE for >= DebounceTime
 * Weld_Soft_Start_Active: TRUE during INIT (PUB005), FALSE otherwise
 *
 * Reset/priority: E_Stop FALSE (active) >> INIT >> MONITOR/ALARM
 * - E_Stop: clears alarm, timers (PUB004)
 * - Gap FALSE: clears alarm, debounce timer (PUB003)
 * - No latching; alarm is level-driven by debounced gap
 *)
VAR_INPUT
    Gap_Exceeded   : BOOL;
    Weld_E_Stop_NC : BOOL;
    DebounceTime   : TIME;
END_VAR

VAR_OUTPUT
    Operator_Alert         : BOOL := FALSE;
    Weld_Soft_Start_Active : BOOL := TRUE;
END_VAR

VAR
    init_timer           : TON;
    debounce_timer       : TON;
    init_complete        : BOOL := FALSE;
    tmp_debounce_started : BOOL := FALSE;
END_VAR

    // E-Stop priority: active when Weld_E_Stop_NC = FALSE
    IF NOT Weld_E_Stop_NC THEN
        Operator_Alert          := FALSE;
        Weld_Soft_Start_Active  := FALSE;
        debounce_timer(IN := FALSE);
        init_timer(IN := FALSE);
        init_complete         := FALSE;
        tmp_debounce_started  := FALSE;
        RETURN;
    END_IF;

    // Normal monitoring: debounce gap signal (PUB003)
    IF init_complete THEN
        Operator_Alert := FALSE;

        IF Gap_Exceeded THEN
            // Start debounce timer only on first TRUE detection
            IF NOT tmp_debounce_started THEN
                debounce_timer(IN := TRUE, PT := DebounceTime);
                tmp_debounce_started := TRUE;
            END_IF;
            Operator_Alert := debounce_timer.Q;
        ELSE
            debounce_timer(IN := FALSE);
            tmp_debounce_started := FALSE;
        END_IF;

    // Initialization: 5-second power-up inhibition (PUB002, PUB005)
    ELSE
        // Keep init timer running continuously while not complete
        init_timer(IN := TRUE, PT := T#5S);
        Weld_Soft_Start_Active := TRUE;
        Operator_Alert         := FALSE;
        debounce_timer(IN := FALSE);

        IF init_timer.Q THEN
            init_complete          := TRUE;
            Weld_Soft_Start_Active := FALSE;
            init_timer(IN := FALSE);
        END_IF;
    END_IF;

END_FUNCTION_BLOCK
(* CONTRACT_RULES [] *)

(* ---- public-easy-05.candidate_03.st ---- *)
FUNCTION_BLOCK Weld_Gap_Alarm
(* ENGINEERING_CONTRACT
 * States: INIT(5s inhibit) | MONITOR(gap OK) | ALARM(gap debounced)
 *
 * Operator_Alert: FALSE during INIT, TRUE only when gap TRUE for >= DebounceTime
 * Weld_Soft_Start_Active: TRUE during INIT (PUB005), FALSE otherwise
 *
 * Reset/priority: E_Stop FALSE (active) >> INIT >> MONITOR/ALARM
 * - E_Stop: clears alarm, timers (PUB004)
 * - Gap FALSE: clears alarm, debounce timer (PUB003)
 * - No latching; alarm is level-driven by debounced gap
 *)
VAR_INPUT
    Gap_Exceeded   : BOOL;
    Weld_E_Stop_NC : BOOL;
    DebounceTime   : TIME;
END_VAR

VAR_OUTPUT
    Operator_Alert         : BOOL := FALSE;
    Weld_Soft_Start_Active : BOOL := TRUE;
END_VAR

VAR
    init_timer     : TON;
    debounce_timer : TON;
    init_complete  : BOOL := FALSE;
END_VAR

    // E-Stop priority: active when Weld_E_Stop_NC = FALSE
    IF NOT Weld_E_Stop_NC THEN
        Operator_Alert         := FALSE;
        Weld_Soft_Start_Active := FALSE;
        debounce_timer(IN := FALSE);
        init_timer(IN := FALSE);
        init_complete := FALSE;
        RETURN;
    END_IF;

    // Initialization: 5-second power-up inhibition (PUB002, PUB005)
    IF NOT init_complete THEN
        init_timer(IN := NOT init_complete, PT := T#5S);
        Weld_Soft_Start_Active := TRUE;
        Operator_Alert         := FALSE;
        debounce_timer(IN := FALSE);

        IF init_timer.Q THEN
            init_complete          := TRUE;
            Weld_Soft_Start_Active := FALSE;
        END_IF;

    // Normal monitoring: debounce gap signal (PUB003)
    ELSE
        Operator_Alert := FALSE;

        IF Gap_Exceeded THEN
            debounce_timer(IN := TRUE, PT := DebounceTime);
            Operator_Alert := debounce_timer.Q;
        ELSE
            debounce_timer(IN := FALSE);
        END_IF;
    END_IF;

END_FUNCTION_BLOCK
(* CONTRACT_RULES [] *)

(* ---- public-easy-05.candidate_04.st ---- *)
FUNCTION_BLOCK Weld_Gap_Alarm
(* ENGINEERING_CONTRACT
 * States: INIT(5s inhibit) | MONITOR(gap OK) | ALARM(gap debounced)
 *
 * Operator_Alert: FALSE during INIT, TRUE only when gap TRUE for >= DebounceTime
 * Weld_Soft_Start_Active: TRUE during INIT (PUB005), FALSE otherwise
 *
 * Reset/priority: E_Stop FALSE (active) >> INIT >> MONITOR/ALARM
 * - E_Stop: clears alarm, timers, init state (PUB004)
 * - Gap FALSE: clears alarm, debounce timer (PUB003)
 * - Init complete: explicit debounce_timer reset prevents ET bleed-through
 * - No latching; alarm is level-driven by debounced gap
 *)
VAR_INPUT
    Gap_Exceeded   : BOOL;
    Weld_E_Stop_NC : BOOL;
    DebounceTime   : TIME;
END_VAR

VAR_OUTPUT
    Operator_Alert         : BOOL := FALSE;
    Weld_Soft_Start_Active : BOOL := TRUE;
END_VAR

VAR
    init_timer     : TON;
    debounce_timer : TON;
    init_complete  : BOOL := FALSE;
END_VAR

    // E-Stop priority: active when Weld_E_Stop_NC = FALSE
    IF NOT Weld_E_Stop_NC THEN
        Operator_Alert         := FALSE;
        Weld_Soft_Start_Active := FALSE;
        debounce_timer(IN := FALSE);
        init_timer(IN := FALSE);
        init_complete := FALSE;
        RETURN;
    END_IF;

    // Initialization: 5-second power-up inhibition (PUB002, PUB005)
    IF NOT init_complete THEN
        init_timer(IN := TRUE, PT := T#5S);
        Weld_Soft_Start_Active := TRUE;
        Operator_Alert         := FALSE;
        debounce_timer(IN := FALSE);

        IF init_timer.Q THEN
            init_complete          := TRUE;
            Weld_Soft_Start_Active := FALSE;
            init_timer(IN := FALSE);
            debounce_timer(IN := FALSE); // Reset to prevent ET bleed-through
        END_IF;

    // Normal monitoring: debounce gap signal (PUB003)
    ELSE
        Operator_Alert := FALSE;

        IF Gap_Exceeded THEN
            debounce_timer(IN := TRUE, PT := DebounceTime);
            Operator_Alert := debounce_timer.Q;
        ELSE
            debounce_timer(IN := FALSE);
        END_IF;
    END_IF;

END_FUNCTION_BLOCK
(* CONTRACT_RULES [] *)

(* ---- public-easy-05.raw_candidate_01.st ---- *)
FUNCTION_BLOCK Weld_Gap_Alarm
(* ENGINEERING_CONTRACT
 * States: INIT(5s inhibit) | MONITOR(gap OK) | ALARM(gap debounced)
 *
 * Operator_Alert: FALSE during INIT, TRUE only when gap TRUE for >= DebounceTime
 * Weld_Soft_Start_Active: TRUE during INIT (PUB005), FALSE otherwise
 *
 * Reset/priority: E_Stop FALSE (active) >> INIT >> MONITOR/ALARM
 * - E_Stop: clears alarm, timers (PUB004)
 * - Gap FALSE: clears alarm, debounce timer (PUB003)
 * - No latching; alarm is level-driven by debounced gap
 *)
VAR_INPUT
    Gap_Exceeded   : BOOL;
    Weld_E_Stop_NC : BOOL;
    DebounceTime   : TIME;
END_VAR

VAR_OUTPUT
    Operator_Alert        : BOOL := FALSE;
    Weld_Soft_Start_Active : BOOL := TRUE;
END_VAR

VAR
    init_timer      : TON;
    debounce_timer  : TON;
    init_complete   : BOOL := FALSE;
END_VAR

    // E-Stop priority: active when Weld_E_Stop_NC = FALSE
    IF NOT Weld_E_Stop_NC THEN
        Operator_Alert         := FALSE;
        Weld_Soft_Start_Active := FALSE;
        debounce_timer(IN := FALSE);
        init_timer(IN := FALSE);
        init_complete := FALSE;
        RETURN;
    END_IF;

    // Initialization: 5-second power-up inhibition (PUB002, PUB005)
    IF NOT init_complete THEN
        init_timer(IN := TRUE, PT := T#5S);
        Weld_Soft_Start_Active := TRUE;
        Operator_Alert         := FALSE;
        debounce_timer(IN := FALSE);

        IF init_timer.Q THEN
            init_complete          := TRUE;
            Weld_Soft_Start_Active := FALSE;
            init_timer(IN := FALSE);
        END_IF;

    // Normal monitoring: debounce gap signal (PUB003)
    ELSE
        Operator_Alert := FALSE;

        IF Gap_Exceeded THEN
            debounce_timer(IN := TRUE, PT := DebounceTime);
            Operator_Alert := debounce_timer.Q;
        ELSE
            debounce_timer(IN := FALSE);
        END_IF;
    END_IF;

END_FUNCTION_BLOCK
(* CONTRACT_RULES [] *)

(* ---- public-easy-05.raw_candidate_02.st ---- *)
FUNCTION_BLOCK Weld_Gap_Alarm
(* ENGINEERING_CONTRACT
 * States: INIT(5s inhibit) | MONITOR(gap OK) | ALARM(gap debounced)
 *
 * Operator_Alert: FALSE during INIT, TRUE only when gap TRUE for >= DebounceTime
 * Weld_Soft_Start_Active: TRUE during INIT (PUB005), FALSE otherwise
 *
 * Reset/priority: E_Stop FALSE (active) >> INIT >> MONITOR/ALARM
 * - E_Stop: clears alarm, timers (PUB004)
 * - Gap FALSE: clears alarm, debounce timer (PUB003)
 * - No latching; alarm is level-driven by debounced gap
 *)
VAR_INPUT
    Gap_Exceeded   : BOOL;
    Weld_E_Stop_NC : BOOL;
    DebounceTime   : TIME;
END_VAR

VAR_OUTPUT
    Operator_Alert         : BOOL := FALSE;
    Weld_Soft_Start_Active : BOOL := TRUE;
END_VAR

VAR
    init_timer           : TON;
    debounce_timer       : TON;
    init_complete        : BOOL := FALSE;
    tmp_debounce_started : BOOL := FALSE;
END_VAR

    // E-Stop priority: active when Weld_E_Stop_NC = FALSE
    IF NOT Weld_E_Stop_NC THEN
        Operator_Alert          := FALSE;
        Weld_Soft_Start_Active  := FALSE;
        debounce_timer(IN := FALSE);
        init_timer(IN := FALSE);
        init_complete         := FALSE;
        tmp_debounce_started  := FALSE;
        RETURN;
    END_IF;

    // Normal monitoring: debounce gap signal (PUB003)
    IF init_complete THEN
        Operator_Alert := FALSE;

        IF Gap_Exceeded THEN
            // Start debounce timer only on first TRUE detection
            IF NOT tmp_debounce_started THEN
                debounce_timer(IN := TRUE, PT := DebounceTime);
                tmp_debounce_started := TRUE;
            END_IF;
            Operator_Alert := debounce_timer.Q;
        ELSE
            debounce_timer(IN := FALSE);
            tmp_debounce_started := FALSE;
        END_IF;

    // Initialization: 5-second power-up inhibition (PUB002, PUB005)
    ELSE
        // Keep init timer running continuously while not complete
        init_timer(IN := TRUE, PT := T#5S);
        Weld_Soft_Start_Active := TRUE;
        Operator_Alert         := FALSE;
        debounce_timer(IN := FALSE);

        IF init_timer.Q THEN
            init_complete          := TRUE;
            Weld_Soft_Start_Active := FALSE;
            init_timer(IN := FALSE);
        END_IF;
    END_IF;

END_FUNCTION_BLOCK
(* CONTRACT_RULES [] *)

(* ---- public-easy-05.raw_candidate_03.st ---- *)
FUNCTION_BLOCK Weld_Gap_Alarm
(* ENGINEERING_CONTRACT
 * States: INIT(5s inhibit) | MONITOR(gap OK) | ALARM(gap debounced)
 *
 * Operator_Alert: FALSE during INIT, TRUE only when gap TRUE for >= DebounceTime
 * Weld_Soft_Start_Active: TRUE during INIT (PUB005), FALSE otherwise
 *
 * Reset/priority: E_Stop FALSE (active) >> INIT >> MONITOR/ALARM
 * - E_Stop: clears alarm, timers (PUB004)
 * - Gap FALSE: clears alarm, debounce timer (PUB003)
 * - No latching; alarm is level-driven by debounced gap
 *)
VAR_INPUT
    Gap_Exceeded   : BOOL;
    Weld_E_Stop_NC : BOOL;
    DebounceTime   : TIME;
END_VAR

VAR_OUTPUT
    Operator_Alert         : BOOL := FALSE;
    Weld_Soft_Start_Active : BOOL := TRUE;
END_VAR

VAR
    init_timer     : TON;
    debounce_timer : TON;
    init_complete  : BOOL := FALSE;
END_VAR

    // E-Stop priority: active when Weld_E_Stop_NC = FALSE
    IF NOT Weld_E_Stop_NC THEN
        Operator_Alert         := FALSE;
        Weld_Soft_Start_Active := FALSE;
        debounce_timer(IN := FALSE);
        init_timer(IN := FALSE);
        init_complete := FALSE;
        RETURN;
    END_IF;

    // Initialization: 5-second power-up inhibition (PUB002, PUB005)
    IF NOT init_complete THEN
        init_timer(IN := NOT init_complete, PT := T#5S);
        Weld_Soft_Start_Active := TRUE;
        Operator_Alert         := FALSE;
        debounce_timer(IN := FALSE);

        IF init_timer.Q THEN
            init_complete          := TRUE;
            Weld_Soft_Start_Active := FALSE;
        END_IF;

    // Normal monitoring: debounce gap signal (PUB003)
    ELSE
        Operator_Alert := FALSE;

        IF Gap_Exceeded THEN
            debounce_timer(IN := TRUE, PT := DebounceTime);
            Operator_Alert := debounce_timer.Q;
        ELSE
            debounce_timer(IN := FALSE);
        END_IF;
    END_IF;

END_FUNCTION_BLOCK
(* CONTRACT_RULES [] *)

(* ---- public-easy-05.raw_candidate_04.st ---- *)
FUNCTION_BLOCK Weld_Gap_Alarm
(* ENGINEERING_CONTRACT
 * States: INIT(5s inhibit) | MONITOR(gap OK) | ALARM(gap debounced)
 *
 * Operator_Alert: FALSE during INIT, TRUE only when gap TRUE for >= DebounceTime
 * Weld_Soft_Start_Active: TRUE during INIT (PUB005), FALSE otherwise
 *
 * Reset/priority: E_Stop FALSE (active) >> INIT >> MONITOR/ALARM
 * - E_Stop: clears alarm, timers, init state (PUB004)
 * - Gap FALSE: clears alarm, debounce timer (PUB003)
 * - Init complete: explicit debounce_timer reset prevents ET bleed-through
 * - No latching; alarm is level-driven by debounced gap
 *)
VAR_INPUT
    Gap_Exceeded   : BOOL;
    Weld_E_Stop_NC : BOOL;
    DebounceTime   : TIME;
END_VAR

VAR_OUTPUT
    Operator_Alert         : BOOL := FALSE;
    Weld_Soft_Start_Active : BOOL := TRUE;
END_VAR

VAR
    init_timer     : TON;
    debounce_timer : TON;
    init_complete  : BOOL := FALSE;
END_VAR

    // E-Stop priority: active when Weld_E_Stop_NC = FALSE
    IF NOT Weld_E_Stop_NC THEN
        Operator_Alert         := FALSE;
        Weld_Soft_Start_Active := FALSE;
        debounce_timer(IN := FALSE);
        init_timer(IN := FALSE);
        init_complete := FALSE;
        RETURN;
    END_IF;

    // Initialization: 5-second power-up inhibition (PUB002, PUB005)
    IF NOT init_complete THEN
        init_timer(IN := TRUE, PT := T#5S);
        Weld_Soft_Start_Active := TRUE;
        Operator_Alert         := FALSE;
        debounce_timer(IN := FALSE);

        IF init_timer.Q THEN
            init_complete          := TRUE;
            Weld_Soft_Start_Active := FALSE;
            init_timer(IN := FALSE);
            debounce_timer(IN := FALSE); // Reset to prevent ET bleed-through
        END_IF;

    // Normal monitoring: debounce gap signal (PUB003)
    ELSE
        Operator_Alert := FALSE;

        IF Gap_Exceeded THEN
            debounce_timer(IN := TRUE, PT := DebounceTime);
            Operator_Alert := debounce_timer.Q;
        ELSE
            debounce_timer(IN := FALSE);
        END_IF;
    END_IF;

END_FUNCTION_BLOCK
(* CONTRACT_RULES [] *)

(* ---- public-easy-06.candidate_01.st ---- *)
(* ENGINEERING_CONTRACT
 * ============================================================
 * PUB001 (81-237): Start delay timing
 *   - Activation: Start TON when DO_LOW AND AERATION_E_STOP_NC both TRUE
 *   - Timer PT: 5 seconds (LTIME, T#5s)
 *   - BLOWER_RUN := TON.Q when timer elapsed
 *   - Retention: BLOWER_RUN held TRUE while conditions remain; no autonomous off
 *
 * PUB002 (239-409): Immediate disable and timer reset
 *   - Deactivation: If DO_LOW = FALSE OR AERATION_E_STOP_NC = FALSE
 *   - BLOWER_RUN := FALSE immediately
 *   - Timer reset (TON.TP.IN := FALSE, TON.ET := 0)
 *   - Must re-wait full 5 seconds on next demand
 *
 * PUB003 (410-614): Cycle count on rising edge
 *   - Set input: BLOWER_RUN rising edge (FALSE->TRUE)
 *   - Increment AERATION_BLOWER_CYCLE_COUNT by 1
 *   - No count during continuous TRUE
 *
 * PUB004 (615-761): Power-up initialization
 *   - BLOWER_RUN := FALSE
 *   - AERATION_BLOWER_CYCLE_COUNT := 0
 *   - Timer state cleared
 *
 * PUB005 (762-910): BOOL enable gate, no speed ramp
 *   - BLOWER_RUN is a simple BOOL command
 *   - No ramp, no intermediate states
 * ============================================================
 *)

(* CONTRACT_RULES [{"kind":"hold_until_reset","output":"BLOWER_RUN","set_input":"internal_timer_done","reset_input":"DO_LOW_OR_ESTOP"}] *)

FUNCTION_BLOCK AerationBlowerDelayedStart
VAR_OUTPUT
    BLOWER_RUN                  : BOOL := FALSE;
    AERATION_BLOWER_CYCLE_COUNT : UINT := 0;
END_VAR
VAR
    StartDelayTimer             : TON;
    BlowerStartRTrig            : R_TRIG;
    ConditionsMet               : BOOL;
    BlowerWasRunning            : BOOL;
END_VAR

// Combine start conditions: DO_LOW AND emergency stop NOT active
ConditionsMet := DO_LOW AND AERATION_E_STOP_NC;

// Start delay timer: enable when conditions met, reset when not
StartDelayTimer(IN := ConditionsMet, PT := T#5s);

// BLOWER_RUN follows timer completion while conditions remain
BLOWER_RUN := StartDelayTimer.Q;

// Rising edge detection on BLOWER_RUN for cycle counting
BlowerStartRTrig(CLK := BLOWER_RUN);
IF BlowerStartRTrig.Q THEN
    AERATION_BLOWER_CYCLE_COUNT := AERATION_BLOWER_CYCLE_COUNT + 1;
END_IF;

END_FUNCTION_BLOCK

(* ---- public-easy-06.candidate_02.st ---- *)
(* ENGINEERING_CONTRACT
 * ============================================================
 * PUB001 (81-237): Start delay timing
 *   - Activation: Start TON when DO_LOW AND AERATION_E_STOP_NC both TRUE
 *   - Timer PT: 5 seconds (LTIME, T#5s)
 *   - BLOWER_RUN := TON.Q when timer elapsed
 *   - Retention: BLOWER_RUN held TRUE while conditions remain; no autonomous off
 *
 * PUB002 (239-409): Immediate disable and timer reset
 *   - Deactivation: If DO_LOW = FALSE OR AERATION_E_STOP_NC = FALSE
 *   - BLOWER_RUN := FALSE immediately
 *   - Timer reset (TON.IN := FALSE, TON.ET := 0)
 *   - Must re-wait full 5 seconds on next demand
 *
 * PUB003 (410-614): Cycle count on rising edge
 *   - Set input: BLOWER_RUN rising edge (FALSE->TRUE)
 *   - Increment AERATION_BLOWER_CYCLE_COUNT by 1
 *   - No count during continuous TRUE
 *
 * PUB004 (615-761): Power-up initialization
 *   - BLOWER_RUN := FALSE
 *   - AERATION_BLOWER_CYCLE_COUNT := 0
 *   - Timer state cleared
 *
 * PUB005 (762-910): BOOL enable gate, no speed ramp
 *   - BLOWER_RUN is a simple BOOL command
 *   - No ramp, no intermediate states
 * ============================================================
 *)

(* CONTRACT_RULES [] *)

FUNCTION_BLOCK AerationBlowerDelayedStart
VAR_INPUT
    DO_LOW                : BOOL;
    AERATION_E_STOP_NC    : BOOL;
END_VAR
VAR_OUTPUT
    BLOWER_RUN                    : BOOL := FALSE;
    AERATION_BLOWER_CYCLE_COUNT   : UINT := 0;
END_VAR
VAR
    StartDelayTimer       : TON;
    BlowerStartRTrig      : R_TRIG;
    tmp_conditions_met    : BOOL;
END_VAR

tmp_conditions_met := DO_LOW AND AERATION_E_STOP_NC;

StartDelayTimer(IN := tmp_conditions_met, PT := T#5s);

BLOWER_RUN := StartDelayTimer.Q;

BlowerStartRTrig(CLK := BLOWER_RUN);
IF BlowerStartRTrig.Q THEN
    AERATION_BLOWER_CYCLE_COUNT := AERATION_BLOWER_CYCLE_COUNT + 1;
END_IF;

END_FUNCTION_BLOCK

(* ---- public-easy-06.raw_candidate_01.st ---- *)
(* ENGINEERING_CONTRACT
 * ============================================================
 * PUB001 (81-237): Start delay timing
 *   - Activation: Start TON when DO_LOW AND AERATION_E_STOP_NC both TRUE
 *   - Timer PT: 5 seconds (LTIME, T#5s)
 *   - BLOWER_RUN := TON.Q when timer elapsed
 *   - Retention: BLOWER_RUN held TRUE while conditions remain; no autonomous off
 *
 * PUB002 (239-409): Immediate disable and timer reset
 *   - Deactivation: If DO_LOW = FALSE OR AERATION_E_STOP_NC = FALSE
 *   - BLOWER_RUN := FALSE immediately
 *   - Timer reset (TON.TP.IN := FALSE, TON.ET := 0)
 *   - Must re-wait full 5 seconds on next demand
 *
 * PUB003 (410-614): Cycle count on rising edge
 *   - Set input: BLOWER_RUN rising edge (FALSE->TRUE)
 *   - Increment AERATION_BLOWER_CYCLE_COUNT by 1
 *   - No count during continuous TRUE
 *
 * PUB004 (615-761): Power-up initialization
 *   - BLOWER_RUN := FALSE
 *   - AERATION_BLOWER_CYCLE_COUNT := 0
 *   - Timer state cleared
 *
 * PUB005 (762-910): BOOL enable gate, no speed ramp
 *   - BLOWER_RUN is a simple BOOL command
 *   - No ramp, no intermediate states
 * ============================================================
 *)

(* CONTRACT_RULES [{"kind":"hold_until_reset","output":"BLOWER_RUN","set_input":"internal_timer_done","reset_input":"DO_LOW_OR_ESTOP"}] *)

FUNCTION_BLOCK AerationBlowerDelayedStart
VAR_OUTPUT
    BLOWER_RUN                  : BOOL := FALSE;
    AERATION_BLOWER_CYCLE_COUNT : UINT := 0;
END_VAR
VAR
    StartDelayTimer             : TON;
    BlowerStartRTrig            : R_TRIG;
    ConditionsMet               : BOOL;
    BlowerWasRunning            : BOOL;
END_VAR

// Combine start conditions: DO_LOW AND emergency stop NOT active
ConditionsMet := DO_LOW AND AERATION_E_STOP_NC;

// Start delay timer: enable when conditions met, reset when not
StartDelayTimer(IN := ConditionsMet, PT := T#5s);

// BLOWER_RUN follows timer completion while conditions remain
BLOWER_RUN := StartDelayTimer.Q;

// Rising edge detection on BLOWER_RUN for cycle counting
BlowerStartRTrig(CLK := BLOWER_RUN);
IF BlowerStartRTrig.Q THEN
    AERATION_BLOWER_CYCLE_COUNT := AERATION_BLOWER_CYCLE_COUNT + 1;
END_IF

END_FUNCTION_BLOCK

(* ---- public-easy-06.raw_candidate_02.st ---- *)
(* ENGINEERING_CONTRACT
 * ============================================================
 * PUB001 (81-237): Start delay timing
 *   - Activation: Start TON when DO_LOW AND AERATION_E_STOP_NC both TRUE
 *   - Timer PT: 5 seconds (LTIME, T#5s)
 *   - BLOWER_RUN := TON.Q when timer elapsed
 *   - Retention: BLOWER_RUN held TRUE while conditions remain; no autonomous off
 *
 * PUB002 (239-409): Immediate disable and timer reset
 *   - Deactivation: If DO_LOW = FALSE OR AERATION_E_STOP_NC = FALSE
 *   - BLOWER_RUN := FALSE immediately
 *   - Timer reset (TON.IN := FALSE, TON.ET := 0)
 *   - Must re-wait full 5 seconds on next demand
 *
 * PUB003 (410-614): Cycle count on rising edge
 *   - Set input: BLOWER_RUN rising edge (FALSE->TRUE)
 *   - Increment AERATION_BLOWER_CYCLE_COUNT by 1
 *   - No count during continuous TRUE
 *
 * PUB004 (615-761): Power-up initialization
 *   - BLOWER_RUN := FALSE
 *   - AERATION_BLOWER_CYCLE_COUNT := 0
 *   - Timer state cleared
 *
 * PUB005 (762-910): BOOL enable gate, no speed ramp
 *   - BLOWER_RUN is a simple BOOL command
 *   - No ramp, no intermediate states
 * ============================================================
 *)

(* CONTRACT_RULES [] *)

FUNCTION_BLOCK AerationBlowerDelayedStart
VAR_INPUT
    DO_LOW                : BOOL;
    AERATION_E_STOP_NC    : BOOL;
END_VAR
VAR_OUTPUT
    BLOWER_RUN                    : BOOL := FALSE;
    AERATION_BLOWER_CYCLE_COUNT   : UINT := 0;
END_VAR
VAR
    StartDelayTimer       : TON;
    BlowerStartRTrig      : R_TRIG;
    tmp_conditions_met    : BOOL;
END_VAR

tmp_conditions_met := DO_LOW AND AERATION_E_STOP_NC;

StartDelayTimer(IN := tmp_conditions_met, PT := T#5s);

BLOWER_RUN := StartDelayTimer.Q;

BlowerStartRTrig(CLK := BLOWER_RUN);
IF BlowerStartRTrig.Q THEN
    AERATION_BLOWER_CYCLE_COUNT := AERATION_BLOWER_CYCLE_COUNT + 1;
END_IF;

END_FUNCTION_BLOCK

(* ---- public-hard-01.candidate_01.st ---- *)
(* ENGINEERING_CONTRACT *)
(*
  PUB001: Emergency stop (estop=FALSE) immediately de-energizes all outputs (valveARun, valveBRun, valveCRun, valveDRun, mixMotorRun).
  PUB002: opeMode=FALSE selects Manual Mode; opeMode=TRUE selects Automatic Mode.
  PUB003: Manual Mode - rising edge on valveAStart toggles valveARun; similarly B/C/D and mixMotorStart each toggle their respective outputs.
  PUB004: Automatic Mode - rising edge on autoStart initiates sequence; valve A opens first.
  PUB005: Level >= 50 cm triggers close valve A + open valve B transition.
  PUB006: Level >= 80 cm triggers close valve B; processMode=FALSE skips valve C; processMode=TRUE proceeds to valve C fill.
  PUB007: processMode=TRUE: valve C opens at level>=80; level>=100 closes valve C.
  PUB008: After level>=80 (or level>=100 for processMode=TRUE), mixing motor starts on mixMotorComplete signal.
  PUB009: mixMotorComplete=TRUE stops mixing motor, opens valve D, and terminates the automatic sequence.
  PUB010: All outputs retain state across scans except when explicitly changed by state transitions or estop.
  PUB011: Rising-edge detection uses R_TRIG on momentary inputs; manual toggles are stateful across scans.
  PUB012: Level sensor thresholds are strict >= comparisons at integer resolution (cm).
  PUB013: No unstated resets, interlocks, or edge triggers beyond R_TRIG on start inputs.
  PUB014: Same-scan priority: output assignments before RETURN; state changes apply to subsequent scan.
  PUB015: Valve/motor stop on estop or mode change takes precedence over automatic sequence state.
*)
(* CONTRACT_RULES [] *)

FUNCTION_BLOCK MaterialProportioning
VAR_INPUT
    estop           : BOOL;
    opeMode         : BOOL;
    valveAStart     : BOOL;
    valveBStart     : BOOL;
    valveCStart     : BOOL;
    valveDStart     : BOOL;
    mixMotorStart   : BOOL;
    autoStart       : BOOL;
    processMode     : BOOL;
    levelSensor     : INT;
    mixMotorComplete: BOOL;
END_VAR
VAR_OUTPUT
    valveARun       : BOOL;
    valveBRun       : BOOL;
    valveCRun       : BOOL;
    valveDRun       : BOOL;
    mixMotorRun     : BOOL;
END_VAR
VAR
    tmp_autoStartTrig    : R_TRIG;
    tmp_valveAStartTrig  : R_TRIG;
    tmp_valveBStartTrig  : R_TRIG;
    tmp_valveCStartTrig  : R_TRIG;
    tmp_valveDStartTrig  : R_TRIG;
    tmp_mixMotorStartTrig: R_TRIG;
    tmp_autoState        : INT;
    tmp_manualValveA     : BOOL;
    tmp_manualValveB     : BOOL;
    tmp_manualValveC     : BOOL;
    tmp_manualValveD     : BOOL;
    tmp_manualMixMotor   : BOOL;
END_VAR

CONSTANTS
    AUTO_IDLE      : INT := 0;
    AUTO_FILL_A    : INT := 1;
    AUTO_FILL_B    : INT := 2;
    AUTO_FILL_C    : INT := 3;
    AUTO_MIXING    : INT := 4;
    AUTO_DRAINING  : INT := 5;
END_CONSTANTS

(* Rising edge detection *)
tmp_autoStartTrig(CLK := autoStart);
tmp_valveAStartTrig(CLK := valveAStart);
tmp_valveBStartTrig(CLK := valveBStart);
tmp_valveCStartTrig(CLK := valveCStart);
tmp_valveDStartTrig(CLK := valveDStart);
tmp_mixMotorStartTrig(CLK := mixMotorStart);

(* Emergency stop: all outputs OFF immediately *)
IF NOT estop THEN
    valveARun  := FALSE;
    valveBRun  := FALSE;
    valveCRun  := FALSE;
    valveDRun  := FALSE;
    mixMotorRun := FALSE;
    tmp_autoState := AUTO_IDLE;
    tmp_manualValveA := FALSE;
    tmp_manualValveB := FALSE;
    tmp_manualValveC := FALSE;
    tmp_manualValveD := FALSE;
    tmp_manualMixMotor := FALSE;
    RETURN;
END_IF;

(* Mode selection *)
IF NOT opeMode THEN
    (* Manual Mode *)
    valveARun  := tmp_manualValveA;
    valveBRun  := tmp_manualValveB;
    valveCRun  := tmp_manualValveC;
    valveDRun  := tmp_manualValveD;
    mixMotorRun := tmp_manualMixMotor;
    tmp_autoState := AUTO_IDLE;

    IF tmp_valveAStartTrig.Q THEN
        tmp_manualValveA := NOT tmp_manualValveA;
    END_IF;
    IF tmp_valveBStartTrig.Q THEN
        tmp_manualValveB := NOT tmp_manualValveB;
    END_IF;
    IF tmp_valveCStartTrig.Q THEN
        tmp_manualValveC := NOT tmp_manualValveC;
    END_IF;
    IF tmp_valveDStartTrig.Q THEN
        tmp_manualValveD := NOT tmp_manualValveD;
    END_IF;
    IF tmp_mixMotorStartTrig.Q THEN
        tmp_manualMixMotor := NOT tmp_manualMixMotor;
    END_IF;
ELSE
    (* Automatic Mode *)
    tmp_manualValveA := FALSE;
    tmp_manualValveB := FALSE;
    tmp_manualValveC := FALSE;
    tmp_manualValveD := FALSE;
    tmp_manualMixMotor := FALSE;

    CASE tmp_autoState OF
        AUTO_IDLE:
            valveARun  := FALSE;
            valveBRun  := FALSE;
            valveCRun  := FALSE;
            valveDRun  := FALSE;
            mixMotorRun := FALSE;
            IF tmp_autoStartTrig.Q THEN
                tmp_autoState := AUTO_FILL_A;
            END_IF;

        AUTO_FILL_A:
            valveARun := TRUE;
            valveBRun := FALSE;
            valveCRun := FALSE;
            valveDRun := FALSE;
            mixMotorRun := FALSE;
            IF levelSensor >= 50 THEN
                valveARun := FALSE;
                valveBRun := TRUE;
                tmp_autoState := AUTO_FILL_B;
            END_IF;

        AUTO_FILL_B:
            valveARun := FALSE;
            valveBRun := TRUE;
            valveCRun := FALSE;
            valveDRun := FALSE;
            mixMotorRun := FALSE;
            IF levelSensor >= 80 THEN
                valveBRun := FALSE;
                IF NOT processMode THEN
                    tmp_autoState := AUTO_MIXING;
                ELSE
                    valveCRun := TRUE;
                    tmp_autoState := AUTO_FILL_C;
                END_IF;
            END_IF;

        AUTO_FILL_C:
            valveARun := FALSE;
            valveBRun := FALSE;
            valveCRun := TRUE;
            valveDRun := FALSE;
            mixMotorRun := FALSE;
            IF levelSensor >= 100 THEN
                valveCRun := FALSE;
                tmp_autoState := AUTO_MIXING;
            END_IF;

        AUTO_MIXING:
            valveARun := FALSE;
            valveBRun := FALSE;
            valveCRun := FALSE;
            valveDRun := FALSE;
            mixMotorRun := TRUE;
            IF mixMotorComplete THEN
                mixMotorRun := FALSE;
                valveDRun := TRUE;
                tmp_autoState := AUTO_DRAINING;
            END_IF;

        AUTO_DRAINING:
            valveARun := FALSE;
            valveBRun := FALSE;
            valveCRun := FALSE;
            valveDRun := TRUE;
            mixMotorRun := FALSE;
            tmp_autoState := AUTO_IDLE;

    END_CASE;
END_IF;

END_FUNCTION_BLOCK

(* ---- public-hard-01.candidate_02.st ---- *)
(* ENGINEERING_CONTRACT *)
(*
  PUB001: Emergency stop (estop=FALSE) immediately de-energizes all outputs (valveARun, valveBRun, valveCRun, valveDRun, mixMotorRun).
  PUB002: opeMode=FALSE selects Manual Mode; opeMode=TRUE selects Automatic Mode.
  PUB003: Manual Mode - rising edge on valveAStart toggles valveARun; similarly B/C/D and mixMotorStart each toggle their respective outputs.
  PUB004: Automatic Mode - rising edge on autoStart initiates sequence; valve A opens first.
  PUB005: Level >= 50 cm triggers close valve A + open valve B transition.
  PUB006: Level >= 80 cm triggers close valve B; processMode=FALSE skips valve C; processMode=TRUE proceeds to valve C fill.
  PUB007: processMode=TRUE: valve C opens at level>=80; level>=100 closes valve C.
  PUB008: After level>=80 (or level>=100 for processMode=TRUE), mixing motor starts on mixMotorComplete signal.
  PUB009: mixMotorComplete=TRUE stops mixing motor, opens valve D, and terminates the automatic sequence.
  PUB010: All outputs retain state across scans except when explicitly changed by state transitions or estop.
  PUB011: Rising-edge detection uses R_TRIG on momentary inputs; manual toggles are stateful across scans.
  PUB012: Level sensor thresholds are strict >= comparisons at integer resolution (cm).
  PUB013: No unstated resets, interlocks, or edge triggers beyond R_TRIG on start inputs.
  PUB014: Same-scan priority: output assignments before RETURN; state changes apply to subsequent scan.
  PUB015: Valve/motor stop on estop or mode change takes precedence over automatic sequence state.
*)
(* CONTRACT_RULES [] *)

TYPE AutoState :
(
    AUTO_IDLE      := 0,
    AUTO_FILL_A    := 1,
    AUTO_FILL_B    := 2,
    AUTO_FILL_C    := 3,
    AUTO_MIXING    := 4,
    AUTO_DRAINING  := 5
);
END_TYPE;

FUNCTION_BLOCK MaterialProportioning
VAR_INPUT
    estop           : BOOL;
    opeMode         : BOOL;
    valveAStart     : BOOL;
    valveBStart     : BOOL;
    valveCStart     : BOOL;
    valveDStart     : BOOL;
    mixMotorStart   : BOOL;
    autoStart       : BOOL;
    processMode     : BOOL;
    levelSensor     : INT;
    mixMotorComplete: BOOL;
END_VAR
VAR_OUTPUT
    valveARun       : BOOL;
    valveBRun       : BOOL;
    valveCRun       : BOOL;
    valveDRun       : BOOL;
    mixMotorRun     : BOOL;
END_VAR
VAR
    tmp_autoStartTrig    : R_TRIG;
    tmp_valveAStartTrig  : R_TRIG;
    tmp_valveBStartTrig  : R_TRIG;
    tmp_valveCStartTrig  : R_TRIG;
    tmp_valveDStartTrig  : R_TRIG;
    tmp_mixMotorStartTrig: R_TRIG;
    tmp_autoState        : AutoState := AUTO_IDLE;
    tmp_manualValveA     : BOOL;
    tmp_manualValveB     : BOOL;
    tmp_manualValveC     : BOOL;
    tmp_manualValveD     : BOOL;
    tmp_manualMixMotor   : BOOL;
END_VAR

(* Rising edge detection *)
tmp_autoStartTrig(CLK := autoStart);
tmp_valveAStartTrig(CLK := valveAStart);
tmp_valveBStartTrig(CLK := valveBStart);
tmp_valveCStartTrig(CLK := valveCStart);
tmp_valveDStartTrig(CLK := valveDStart);
tmp_mixMotorStartTrig(CLK := mixMotorStart);

(* Emergency stop: all outputs OFF immediately *)
IF NOT estop THEN
    valveARun  := FALSE;
    valveBRun  := FALSE;
    valveCRun  := FALSE;
    valveDRun  := FALSE;
    mixMotorRun := FALSE;
    tmp_autoState := AUTO_IDLE;
    tmp_manualValveA := FALSE;
    tmp_manualValveB := FALSE;
    tmp_manualValveC := FALSE;
    tmp_manualValveD := FALSE;
    tmp_manualMixMotor := FALSE;
    RETURN;
END_IF;

(* Mode selection *)
IF NOT opeMode THEN
    (* Manual Mode *)
    valveARun  := tmp_manualValveA;
    valveBRun  := tmp_manualValveB;
    valveCRun  := tmp_manualValveC;
    valveDRun  := tmp_manualValveD;
    mixMotorRun := tmp_manualMixMotor;
    tmp_autoState := AUTO_IDLE;

    IF tmp_valveAStartTrig.Q THEN
        tmp_manualValveA := NOT tmp_manualValveA;
    END_IF;
    IF tmp_valveBStartTrig.Q THEN
        tmp_manualValveB := NOT tmp_manualValveB;
    END_IF;
    IF tmp_valveCStartTrig.Q THEN
        tmp_manualValveC := NOT tmp_manualValveC;
    END_IF;
    IF tmp_valveDStartTrig.Q THEN
        tmp_manualValveD := NOT tmp_manualValveD;
    END_IF;
    IF tmp_mixMotorStartTrig.Q THEN
        tmp_manualMixMotor := NOT tmp_manualMixMotor;
    END_IF;
ELSE
    (* Automatic Mode *)
    tmp_manualValveA := FALSE;
    tmp_manualValveB := FALSE;
    tmp_manualValveC := FALSE;
    tmp_manualValveD := FALSE;
    tmp_manualMixMotor := FALSE;

    CASE TO_INT(tmp_autoState) OF
        0: (* AUTO_IDLE *)
            valveARun  := FALSE;
            valveBRun  := FALSE;
            valveCRun  := FALSE;
            valveDRun  := FALSE;
            mixMotorRun := FALSE;
            IF tmp_autoStartTrig.Q THEN
                tmp_autoState := AUTO_FILL_A;
            END_IF;

        1: (* AUTO_FILL_A *)
            valveARun := TRUE;
            valveBRun := FALSE;
            valveCRun := FALSE;
            valveDRun := FALSE;
            mixMotorRun := FALSE;
            IF levelSensor >= 50 THEN
                valveARun := FALSE;
                valveBRun := TRUE;
                tmp_autoState := AUTO_FILL_B;
            END_IF;

        2: (* AUTO_FILL_B *)
            valveARun := FALSE;
            valveBRun := TRUE;
            valveCRun := FALSE;
            valveDRun := FALSE;
            mixMotorRun := FALSE;
            IF levelSensor >= 80 THEN
                valveBRun := FALSE;
                IF NOT processMode THEN
                    tmp_autoState := AUTO_MIXING;
                ELSE
                    valveCRun := TRUE;
                    tmp_autoState := AUTO_FILL_C;
                END_IF;
            END_IF;

        3: (* AUTO_FILL_C *)
            valveARun := FALSE;
            valveBRun := FALSE;
            valveCRun := TRUE;
            valveDRun := FALSE;
            mixMotorRun := FALSE;
            IF levelSensor >= 100 THEN
                valveCRun := FALSE;
                tmp_autoState := AUTO_MIXING;
            END_IF;

        4: (* AUTO_MIXING *)
            valveARun := FALSE;
            valveBRun := FALSE;
            valveCRun := FALSE;
            valveDRun := FALSE;
            mixMotorRun := TRUE;
            IF mixMotorComplete THEN
                mixMotorRun := FALSE;
                valveDRun := TRUE;
                tmp_autoState := AUTO_DRAINING;
            END_IF;

        5: (* AUTO_DRAINING *)
            valveARun := FALSE;
            valveBRun := FALSE;
            valveCRun := FALSE;
            valveDRun := TRUE;
            mixMotorRun := FALSE;
            tmp_autoState := AUTO_IDLE;

    END_CASE;
END_IF;

END_FUNCTION_BLOCK

(* ---- public-hard-01.raw_candidate_01.st ---- *)
(* ENGINEERING_CONTRACT *)
(*
  PUB001: Emergency stop (estop=FALSE) immediately de-energizes all outputs (valveARun, valveBRun, valveCRun, valveDRun, mixMotorRun).
  PUB002: opeMode=FALSE selects Manual Mode; opeMode=TRUE selects Automatic Mode.
  PUB003: Manual Mode - rising edge on valveAStart toggles valveARun; similarly B/C/D and mixMotorStart each toggle their respective outputs.
  PUB004: Automatic Mode - rising edge on autoStart initiates sequence; valve A opens first.
  PUB005: Level >= 50 cm triggers close valve A + open valve B transition.
  PUB006: Level >= 80 cm triggers close valve B; processMode=FALSE skips valve C; processMode=TRUE proceeds to valve C fill.
  PUB007: processMode=TRUE: valve C opens at level>=80; level>=100 closes valve C.
  PUB008: After level>=80 (or level>=100 for processMode=TRUE), mixing motor starts on mixMotorComplete signal.
  PUB009: mixMotorComplete=TRUE stops mixing motor, opens valve D, and terminates the automatic sequence.
  PUB010: All outputs retain state across scans except when explicitly changed by state transitions or estop.
  PUB011: Rising-edge detection uses R_TRIG on momentary inputs; manual toggles are stateful across scans.
  PUB012: Level sensor thresholds are strict >= comparisons at integer resolution (cm).
  PUB013: No unstated resets, interlocks, or edge triggers beyond R_TRIG on start inputs.
  PUB014: Same-scan priority: output assignments before RETURN; state changes apply to subsequent scan.
  PUB015: Valve/motor stop on estop or mode change takes precedence over automatic sequence state.
*)
(* CONTRACT_RULES [] *)

FUNCTION_BLOCK MaterialProportioning
VAR_INPUT
    estop           : BOOL;
    opeMode         : BOOL;
    valveAStart     : BOOL;
    valveBStart     : BOOL;
    valveCStart     : BOOL;
    valveDStart     : BOOL;
    mixMotorStart   : BOOL;
    autoStart       : BOOL;
    processMode     : BOOL;
    levelSensor     : INT;
    mixMotorComplete: BOOL;
END_VAR
VAR_OUTPUT
    valveARun       : BOOL;
    valveBRun       : BOOL;
    valveCRun       : BOOL;
    valveDRun       : BOOL;
    mixMotorRun     : BOOL;
END_VAR
VAR
    tmp_autoStartTrig    : R_TRIG;
    tmp_valveAStartTrig  : R_TRIG;
    tmp_valveBStartTrig  : R_TRIG;
    tmp_valveCStartTrig  : R_TRIG;
    tmp_valveDStartTrig  : R_TRIG;
    tmp_mixMotorStartTrig: R_TRIG;
    tmp_autoState        : INT;
    tmp_manualValveA     : BOOL;
    tmp_manualValveB     : BOOL;
    tmp_manualValveC     : BOOL;
    tmp_manualValveD     : BOOL;
    tmp_manualMixMotor   : BOOL;
END_VAR

CONSTANTS
    AUTO_IDLE      : INT := 0;
    AUTO_FILL_A    : INT := 1;
    AUTO_FILL_B    : INT := 2;
    AUTO_FILL_C    : INT := 3;
    AUTO_MIXING    : INT := 4;
    AUTO_DRAINING  : INT := 5;
END_CONSTANTS

(* Rising edge detection *)
tmp_autoStartTrig(CLK := autoStart);
tmp_valveAStartTrig(CLK := valveAStart);
tmp_valveBStartTrig(CLK := valveBStart);
tmp_valveCStartTrig(CLK := valveCStart);
tmp_valveDStartTrig(CLK := valveDStart);
tmp_mixMotorStartTrig(CLK := mixMotorStart);

(* Emergency stop: all outputs OFF immediately *)
IF NOT estop THEN
    valveARun  := FALSE;
    valveBRun  := FALSE;
    valveCRun  := FALSE;
    valveDRun  := FALSE;
    mixMotorRun := FALSE;
    tmp_autoState := AUTO_IDLE;
    tmp_manualValveA := FALSE;
    tmp_manualValveB := FALSE;
    tmp_manualValveC := FALSE;
    tmp_manualValveD := FALSE;
    tmp_manualMixMotor := FALSE;
    RETURN;
END_IF

(* Mode selection *)
IF NOT opeMode THEN
    (* Manual Mode *)
    valveARun  := tmp_manualValveA;
    valveBRun  := tmp_manualValveB;
    valveCRun  := tmp_manualValveC;
    valveDRun  := tmp_manualValveD;
    mixMotorRun := tmp_manualMixMotor;
    tmp_autoState := AUTO_IDLE;

    IF tmp_valveAStartTrig.Q THEN
        tmp_manualValveA := NOT tmp_manualValveA;
    END_IF
    IF tmp_valveBStartTrig.Q THEN
        tmp_manualValveB := NOT tmp_manualValveB;
    END_IF
    IF tmp_valveCStartTrig.Q THEN
        tmp_manualValveC := NOT tmp_manualValveC;
    END_IF
    IF tmp_valveDStartTrig.Q THEN
        tmp_manualValveD := NOT tmp_manualValveD;
    END_IF
    IF tmp_mixMotorStartTrig.Q THEN
        tmp_manualMixMotor := NOT tmp_manualMixMotor;
    END_IF;
ELSE
    (* Automatic Mode *)
    tmp_manualValveA := FALSE;
    tmp_manualValveB := FALSE;
    tmp_manualValveC := FALSE;
    tmp_manualValveD := FALSE;
    tmp_manualMixMotor := FALSE;

    CASE tmp_autoState OF
        AUTO_IDLE:
            valveARun  := FALSE;
            valveBRun  := FALSE;
            valveCRun  := FALSE;
            valveDRun  := FALSE;
            mixMotorRun := FALSE;
            IF tmp_autoStartTrig.Q THEN
                tmp_autoState := AUTO_FILL_A;
            END_IF;

        AUTO_FILL_A:
            valveARun := TRUE;
            valveBRun := FALSE;
            valveCRun := FALSE;
            valveDRun := FALSE;
            mixMotorRun := FALSE;
            IF levelSensor >= 50 THEN
                valveARun := FALSE;
                valveBRun := TRUE;
                tmp_autoState := AUTO_FILL_B;
            END_IF;

        AUTO_FILL_B:
            valveARun := FALSE;
            valveBRun := TRUE;
            valveCRun := FALSE;
            valveDRun := FALSE;
            mixMotorRun := FALSE;
            IF levelSensor >= 80 THEN
                valveBRun := FALSE;
                IF NOT processMode THEN
                    tmp_autoState := AUTO_MIXING;
                ELSE
                    valveCRun := TRUE;
                    tmp_autoState := AUTO_FILL_C;
                END_IF;
            END_IF;

        AUTO_FILL_C:
            valveARun := FALSE;
            valveBRun := FALSE;
            valveCRun := TRUE;
            valveDRun := FALSE;
            mixMotorRun := FALSE;
            IF levelSensor >= 100 THEN
                valveCRun := FALSE;
                tmp_autoState := AUTO_MIXING;
            END_IF;

        AUTO_MIXING:
            valveARun := FALSE;
            valveBRun := FALSE;
            valveCRun := FALSE;
            valveDRun := FALSE;
            mixMotorRun := TRUE;
            IF mixMotorComplete THEN
                mixMotorRun := FALSE;
                valveDRun := TRUE;
                tmp_autoState := AUTO_DRAINING;
            END_IF;

        AUTO_DRAINING:
            valveARun := FALSE;
            valveBRun := FALSE;
            valveCRun := FALSE;
            valveDRun := TRUE;
            mixMotorRun := FALSE;
            tmp_autoState := AUTO_IDLE;

    END_CASE;
END_IF;

END_FUNCTION_BLOCK

(* ---- public-hard-01.raw_candidate_02.st ---- *)
(* ENGINEERING_CONTRACT *)
(*
  PUB001: Emergency stop (estop=FALSE) immediately de-energizes all outputs (valveARun, valveBRun, valveCRun, valveDRun, mixMotorRun).
  PUB002: opeMode=FALSE selects Manual Mode; opeMode=TRUE selects Automatic Mode.
  PUB003: Manual Mode - rising edge on valveAStart toggles valveARun; similarly B/C/D and mixMotorStart each toggle their respective outputs.
  PUB004: Automatic Mode - rising edge on autoStart initiates sequence; valve A opens first.
  PUB005: Level >= 50 cm triggers close valve A + open valve B transition.
  PUB006: Level >= 80 cm triggers close valve B; processMode=FALSE skips valve C; processMode=TRUE proceeds to valve C fill.
  PUB007: processMode=TRUE: valve C opens at level>=80; level>=100 closes valve C.
  PUB008: After level>=80 (or level>=100 for processMode=TRUE), mixing motor starts on mixMotorComplete signal.
  PUB009: mixMotorComplete=TRUE stops mixing motor, opens valve D, and terminates the automatic sequence.
  PUB010: All outputs retain state across scans except when explicitly changed by state transitions or estop.
  PUB011: Rising-edge detection uses R_TRIG on momentary inputs; manual toggles are stateful across scans.
  PUB012: Level sensor thresholds are strict >= comparisons at integer resolution (cm).
  PUB013: No unstated resets, interlocks, or edge triggers beyond R_TRIG on start inputs.
  PUB014: Same-scan priority: output assignments before RETURN; state changes apply to subsequent scan.
  PUB015: Valve/motor stop on estop or mode change takes precedence over automatic sequence state.
*)
(* CONTRACT_RULES [] *)

TYPE AutoState :
(
    AUTO_IDLE      := 0,
    AUTO_FILL_A    := 1,
    AUTO_FILL_B    := 2,
    AUTO_FILL_C    := 3,
    AUTO_MIXING    := 4,
    AUTO_DRAINING  := 5
);
END_TYPE

FUNCTION_BLOCK MaterialProportioning
VAR_INPUT
    estop           : BOOL;
    opeMode         : BOOL;
    valveAStart     : BOOL;
    valveBStart     : BOOL;
    valveCStart     : BOOL;
    valveDStart     : BOOL;
    mixMotorStart   : BOOL;
    autoStart       : BOOL;
    processMode     : BOOL;
    levelSensor     : INT;
    mixMotorComplete: BOOL;
END_VAR
VAR_OUTPUT
    valveARun       : BOOL;
    valveBRun       : BOOL;
    valveCRun       : BOOL;
    valveDRun       : BOOL;
    mixMotorRun     : BOOL;
END_VAR
VAR
    tmp_autoStartTrig    : R_TRIG;
    tmp_valveAStartTrig  : R_TRIG;
    tmp_valveBStartTrig  : R_TRIG;
    tmp_valveCStartTrig  : R_TRIG;
    tmp_valveDStartTrig  : R_TRIG;
    tmp_mixMotorStartTrig: R_TRIG;
    tmp_autoState        : AutoState := AUTO_IDLE;
    tmp_manualValveA     : BOOL;
    tmp_manualValveB     : BOOL;
    tmp_manualValveC     : BOOL;
    tmp_manualValveD     : BOOL;
    tmp_manualMixMotor   : BOOL;
END_VAR

(* Rising edge detection *)
tmp_autoStartTrig(CLK := autoStart);
tmp_valveAStartTrig(CLK := valveAStart);
tmp_valveBStartTrig(CLK := valveBStart);
tmp_valveCStartTrig(CLK := valveCStart);
tmp_valveDStartTrig(CLK := valveDStart);
tmp_mixMotorStartTrig(CLK := mixMotorStart);

(* Emergency stop: all outputs OFF immediately *)
IF NOT estop THEN
    valveARun  := FALSE;
    valveBRun  := FALSE;
    valveCRun  := FALSE;
    valveDRun  := FALSE;
    mixMotorRun := FALSE;
    tmp_autoState := AUTO_IDLE;
    tmp_manualValveA := FALSE;
    tmp_manualValveB := FALSE;
    tmp_manualValveC := FALSE;
    tmp_manualValveD := FALSE;
    tmp_manualMixMotor := FALSE;
    RETURN;
END_IF;

(* Mode selection *)
IF NOT opeMode THEN
    (* Manual Mode *)
    valveARun  := tmp_manualValveA;
    valveBRun  := tmp_manualValveB;
    valveCRun  := tmp_manualValveC;
    valveDRun  := tmp_manualValveD;
    mixMotorRun := tmp_manualMixMotor;
    tmp_autoState := AUTO_IDLE;

    IF tmp_valveAStartTrig.Q THEN
        tmp_manualValveA := NOT tmp_manualValveA;
    END_IF;
    IF tmp_valveBStartTrig.Q THEN
        tmp_manualValveB := NOT tmp_manualValveB;
    END_IF;
    IF tmp_valveCStartTrig.Q THEN
        tmp_manualValveC := NOT tmp_manualValveC;
    END_IF;
    IF tmp_valveDStartTrig.Q THEN
        tmp_manualValveD := NOT tmp_manualValveD;
    END_IF;
    IF tmp_mixMotorStartTrig.Q THEN
        tmp_manualMixMotor := NOT tmp_manualMixMotor;
    END_IF;
ELSE
    (* Automatic Mode *)
    tmp_manualValveA := FALSE;
    tmp_manualValveB := FALSE;
    tmp_manualValveC := FALSE;
    tmp_manualValveD := FALSE;
    tmp_manualMixMotor := FALSE;

    CASE TO_INT(tmp_autoState) OF
        0: (* AUTO_IDLE *)
            valveARun  := FALSE;
            valveBRun  := FALSE;
            valveCRun  := FALSE;
            valveDRun  := FALSE;
            mixMotorRun := FALSE;
            IF tmp_autoStartTrig.Q THEN
                tmp_autoState := AUTO_FILL_A;
            END_IF;

        1: (* AUTO_FILL_A *)
            valveARun := TRUE;
            valveBRun := FALSE;
            valveCRun := FALSE;
            valveDRun := FALSE;
            mixMotorRun := FALSE;
            IF levelSensor >= 50 THEN
                valveARun := FALSE;
                valveBRun := TRUE;
                tmp_autoState := AUTO_FILL_B;
            END_IF;

        2: (* AUTO_FILL_B *)
            valveARun := FALSE;
            valveBRun := TRUE;
            valveCRun := FALSE;
            valveDRun := FALSE;
            mixMotorRun := FALSE;
            IF levelSensor >= 80 THEN
                valveBRun := FALSE;
                IF NOT processMode THEN
                    tmp_autoState := AUTO_MIXING;
                ELSE
                    valveCRun := TRUE;
                    tmp_autoState := AUTO_FILL_C;
                END_IF;
            END_IF;

        3: (* AUTO_FILL_C *)
            valveARun := FALSE;
            valveBRun := FALSE;
            valveCRun := TRUE;
            valveDRun := FALSE;
            mixMotorRun := FALSE;
            IF levelSensor >= 100 THEN
                valveCRun := FALSE;
                tmp_autoState := AUTO_MIXING;
            END_IF;

        4: (* AUTO_MIXING *)
            valveARun := FALSE;
            valveBRun := FALSE;
            valveCRun := FALSE;
            valveDRun := FALSE;
            mixMotorRun := TRUE;
            IF mixMotorComplete THEN
                mixMotorRun := FALSE;
                valveDRun := TRUE;
                tmp_autoState := AUTO_DRAINING;
            END_IF;

        5: (* AUTO_DRAINING *)
            valveARun := FALSE;
            valveBRun := FALSE;
            valveCRun := FALSE;
            valveDRun := TRUE;
            mixMotorRun := FALSE;
            tmp_autoState := AUTO_IDLE;

    END_CASE;
END_IF;

END_FUNCTION_BLOCK
